(* IEC 61131-3 sources: SortJet_MasterSPS_Aufbau.fbsproj/09_Station/Stationen/_Basic/Aktionen, 11 files *)

(* ---- Basic_Shuttle_Aktion_FB_V01_00_00.fb.st ---- *)
(* METADATA
{
	"v3Meta": {
		"objectGuid": "f063b21c-ee9e-4ece-bc3c-2deffdcf07f3"
	}
}
*)
FUNCTION_BLOCK Basic_Shuttle_Aktion_FB_V01_00_00
VAR_IN_OUT

  // STRUKT
  BasisStationsParameter : StationBasisParameter_ST;

END_VAR
VAR_OUTPUT

  // BOOL
  bprtScheibe : BOOL;

END_VAR
VAR_INPUT

  // BOOL
  bpGeblaeseAktiv        : BOOL;
  bpAutomatikAktiv       : BOOL;
  bpVorAbAuftragAktiv    : BOOL;
  bpZielPositionErreicht : BOOL;

  // WORD
  wWand : WORD;

  // Bausteine
  Glastransport   : REFERENCE TO Shuttle_Glastransport_FB_V01_00_00;
  Kippen          : REFERENCE TO Shuttle_Kippen_V01_00_00;
  Wandverstellung : REFERENCE TO Dickenverstellung_FB_V01_00_00;
  Geblaese        : REFERENCE TO Geblaese_Schuetz_FB_V01_00_00;

END_VAR
VAR

  // Steps_TE
  steplAktion : STEPS_TE;

END_VAR
;
END_FUNCTION_BLOCK

(* ---- Basic_Station_Abnehmen_FB_V01_00_00.fb.st ---- *)
(* METADATA
{
	"v3Meta": {
		"objectGuid": "660d4460-1ddc-44b5-9e6a-0f9c596d74b5"
	}
}
*)
FUNCTION_BLOCK Basic_Station_Abnehmen_FB_V01_00_00 EXTENDS Basic_Station_Aktion_FB_V01_00_00
(* Hinweis:
   - Abnehmen: Station kippt, der Bediener nimmt die Scheiben ab und quittiert jede einzelne
   - Die Aktion schreibt nichts in den Glastransport
   - Kippen nur mit der Ausbaustufe bKippen
*)
VAR_INPUT

  // BOOLEAN
  bpFreigabeErhalten        : BOOL; // Station: Freigabe Si-Kreis (verzoegert) liegt an
  bpGlasAbgenommenQuittiert : BOOL; // Station: Bediener quittiert, dass die Scheibe abgenommen wurde (Taster oder Fusstaster gedrueckt)

  // Bausteine
  Kippen : REFERENCE TO Kippen_FB_V01_00_00;

END_VAR
VAR_OUTPUT

  // BOOLEAN
  bpAbnehmenLampe        : BOOL; // Ampel gruen
  bpSignalScheibeAbnehmen : BOOL; // Taster Scheibe abnehmen (blinkt)
  bpSignalGlasbruch      : BOOL;

END_VAR
VAR

  // INT
  ilScheibenZaehler : INT; // Anzahl der Scheiben, die noch abzunehmen sind

END_VAR
//-------------------------------------------------------------------------------------------------
// ABNEHMEN
//-------------------------------------------------------------------------------------------------
IF ( BasisStationsParameter.bAbnehmen
     AND bpAutomatikAktiv )
THEN
  (* Fehlerbehandlung:
     - Kippen
  *)
  IF ( Kippen.bpFehler ) THEN
    Kippen.bpPositionieren := FALSE;
    BasisStationsParameter.wFehlerNummer := Kippen.wpFehlerNr;
    steplAktion := STEP_900_E;
  END_IF

  CASE steplAktion OF
    // ABNEHMEN =====================
    STEP_0_E:
      (* Hinweis:
         - Freigabe durch Quittierten Si-Kreis da ?
      *)
      bpFehler := FALSE;
      bpSignalScheibeAbnehmen := FALSE;
      BasisStationsParameter.bAbnehmenAbgeschlossen := FALSE;

      IF ( bpFreigabeErhalten ) THEN
        ilScheibenZaehler := WORD_TO_INT( BasisStationsParameter.pAuftrag[cWAND_1].wAnzahlScheiben );
        steplAktion := STEP_10_E;
      END_IF

    // ABNEHMEN =====================
    STEP_10_E:
      (* Hinweis:
         - Pruefen ob das Geblase aktiv ist
           => Sicherung nicht ausgeloest
      *)
      IF ( bpGeblaeseFehler ) THEN
        bpDrosselklappeOeffnen := FALSE;
        BasisStationsParameter.wFehlerNummer := cMELDUNG_ANTRIEB_GEBLAESE;
        steplAktion := STEP_900_E;

      ELSE
        bpDrosselklappeOeffnen := TRUE;
        steplAktion := STEP_20_E;

      END_IF

    // ABNEHMEN =====================
    STEP_20_E:
      IF ( NOT Kippen.bpFehler ) THEN
        bpDrosselklappeOeffnen := TRUE;

        Kippen.epZielPosition := eKippen_Position_84Grad;
        Kippen.bpPositionieren := TRUE;

        steplAktion := STEP_30_E;
      ELSE
        Kippen.bpPositionieren := FALSE;
        BasisStationsParameter.wFehlerNummer := Kippen.wpFehlerNr;
        steplAktion := STEP_900_E;
      END_IF

    // ABNEHMEN =====================
    STEP_30_E:
      IF ( Kippen.bpDone OR NOT BasisStationsParameter.stMKs.stStationsAufbau.bKippen[cWAND_1] ) THEN
        bpDrosselklappeOeffnen := FALSE;
        Kippen.bpPositionieren := FALSE;

        bpAbnehmenLampe         := TRUE;
        bpSignalScheibeAbnehmen := TRUE;

        steplAktion := STEP_50_E;
      END_IF

    // ABNEHMEN =====================
    STEP_50_E:
      bpAbnehmenLampe         := gbFlashbit05sec;
      bpSignalScheibeAbnehmen := gbFlashbit05sec;

      (* Hinweis:
         - Erst die Lichtschranke unterbrechen und zur Station gehen
      *)
      IF ( bpFreigabeErhalten ) THEN
        steplAktion := STEP_60_E;
      END_IF

    // ABNEHMEN =====================
    STEP_60_E:
      bpAbnehmenLampe         := gbFlashbit05sec;
      bpSignalScheibeAbnehmen := gbFlashbit05sec;

      IF ( bpGlasAbgenommenQuittiert ) THEN
        ilScheibenZaehler := ( ilScheibenZaehler - 1 );

        IF ( ilScheibenZaehler > 0 ) THEN
          steplAktion := STEP_70_E;

        ELSE
          bpSignalGlasbruch       := FALSE;
          bpAbnehmenLampe         := FALSE;
          bpSignalScheibeAbnehmen := FALSE;

          steplAktion := STEP_1000_E;
        END_IF
      END_IF

    // ABNEHMEN =====================
    STEP_70_E:
      bpSignalGlasbruch := FALSE;

      IF ( NOT bpGlasAbgenommenQuittiert ) THEN
        steplAktion := STEP_60_E;
      END_IF

    // ABNEHMEN =====================
    STEP_900_E:
      bpFehler := TRUE;
      BasisStationsParameter.bFehler := TRUE;
      Kippen.bpPositionieren := FALSE;

    // ABNEHMEN =====================
    STEP_1000_E:
      BasisStationsParameter.bAbnehmenAbgeschlossen := TRUE;

  // ABNEHMEN =====================
  END_CASE
ELSE
  IF ( steplAktion > STEP_0_E ) THEN
    bpFehler                := FALSE;
    bpDrosselklappeOeffnen  := FALSE;
    bpSignalScheibeAbnehmen := FALSE;
    bpAbnehmenLampe         := FALSE;
    bpSignalGlasbruch       := FALSE;

    Kippen.bpPositionieren  := FALSE;

    BasisStationsParameter.bAbnehmenAbgeschlossen := FALSE;

    steplAktion := STEP_0_E;
  END_IF
END_IF
END_FUNCTION_BLOCK

(* ---- Basic_Station_Aktion_FB_V01_00_00.fb.st ---- *)
(* METADATA
{
	"v3Meta": {
		"objectGuid": "12c9ac0e-b17a-4793-9910-dd4830696017"
	}
}
*)
FUNCTION_BLOCK Basic_Station_Aktion_FB_V01_00_00
(* Hinweis:
   - Basis der wandweisen Aktionen einer Station (Ein-, Aus-, Durch-, Vortransport, Messkopplung)
   - Je Wand eine Instanz, die Station ruft sie in einer Schleife ueber die Waende auf
   - Die Komponenten (Kippen, Hub, Verstellungen ...) gibt es je Station nur einmal; die abgeleiteten
     Bausteine bekommen sie als Referenz
*)
VAR_IN_OUT

  // STRUKT
  BasisStationsParameter : StationBasisParameter_ST;

END_VAR
VAR_OUTPUT

  // BOOL
  bpFehler : BOOL; // Status: Schrittkette steht im Fehler
  bpDrosselklappeOeffnen : BOOL; // Anforderung an die Station: Drosselklappe oeffnen, solange der Transport laeuft (die Station entscheidet ueber den Ausgang)

END_VAR
VAR_INPUT

  // BOOL
  bpAutomatikAktiv       : BOOL;
  bpGeblaeseAktiv        : BOOL;
  bpGeblaeseFehler       : BOOL; // Station: Motorschutz des Geblaeses ausgeloest (Station ohne Geblaese-Baustein)
  bpZielPositionErreicht : BOOL;

  // WORD
  wWand : WORD;

  // Bausteine
  Glastransport : REFERENCE TO Basic_Glastransport_FB_V01_00_00;

END_VAR
VAR

  // Steps_TE
  steplAktion : STEPS_TE;

END_VAR
;
END_FUNCTION_BLOCK

(* ---- Basic_Station_Anlegen_FB_V01_00_00.fb.st ---- *)
(* METADATA
{
	"v3Meta": {
		"objectGuid": "7cf149bd-d1d2-4190-82d5-7daf21613ba4"
	}
}
*)
FUNCTION_BLOCK Basic_Station_Anlegen_FB_V01_00_00 EXTENDS Basic_Station_Aktion_FB_V01_00_00
(* Hinweis:
   - Anlegen von Hand: Die Hoehenkontrolle faehrt auf Position, ggf. Hubrahmen einfahren und Anschlaege ausfahren,
     dann wartet die Aktion auf die Quittierung des Bedieners (Taster / Fusstaster)
   - Die Aktion schreibt nichts in den Glastransport und liest nur die Sensoren
   - Ob angelegt oder eingetragen wird, entscheidet das MMI ueber die Transferstation des Auftrags
     (Transferstation 1 = eigene Station: Anlegen, Fremdanlage: Eintransport; Anlegetisch hinter einer Brechanlage)
   - Mit der VSG-Schnittstelle entscheidet die Station selbst: die Station (Eintransport Schneidlinie) uebernimmt ueber
     bpUebernahmeEintransport oder beendet das Anlegen ueber bpBetriebBeendet
   - Hubrahmen und Anschlag nur mit den Ausbaustufen bHubrahmen und bAnschlag, sonst muessen sie nicht uebergeben werden
*)
VAR_IN_OUT

  // BOOLEAN
  blAnlegenErzwingen : BOOL; // Anlegen wurde erzwungen, die Aktion nimmt die Anforderung entgegen

END_VAR
VAR_INPUT

  // BOOLEAN
  bpAnlegenQuittiert          : BOOL;        // Bediener hat angelegt (steigende Flanke Taster / Fusstaster)
  bpVoraussetzungErfuellt     : BOOL := TRUE; // Station: Voraussetzung zum Start (z.B. Kipparme frei)
  bpAnschlagAutomatischFahren : BOOL;        // Station: Anschlaege fahren automatisch aus
  bpNeustart                  : BOOL;        // Station: Anlegen von vorne beginnen (z.B. nach Umschalten der Anschlaege)
  bpUebernahmeEintransport    : BOOL;        // Station (VSG-Schnittstelle): Eintransport der Schneidlinie uebernimmt, das Anlegen gibt ab
  bpBetriebBeendet            : BOOL;        // Station (VSG-Schnittstelle): Automatikbetrieb der Schneidlinie beendet, Scheibe muss neu angelegt werden

  // Bausteine
  Messachse : REFERENCE TO Messachse_FB_V01_00_00;
  Anschlag  : REFERENCE TO ZylinderPneumatik_Anschlag_FB_V01_00_00;
  Hubrahmen : REFERENCE TO ZylinderPneumatik_Riemen_FB_V01_00_00;

END_VAR
VAR_OUTPUT

  // BOOLEAN
  bpAnlegenLampe          : BOOL; // Ampel gruen / Signal Scheibe aufgegeben (blinkt, bis angelegt ist)
  bpBedienerEingriff      : BOOL; // Aktion wartet auf den Bediener, Handfunktionen (Knebel, Hubrahmen) muessen im Automatikbetrieb greifen
  bpAnlegenInVorbereitung : BOOL; // Aktion fuehrt die Vorbereitung durch (vor dem Warten auf den Bediener)
  bpAnlegenAktiv          : BOOL; // Aktion ist gestartet und noch nicht abgeschlossen
  bpAnlegenFertig         : BOOL; // Aktion hat selbst abgeschlossen (epTypeHoehenmessung gueltig)
  bpGeblaeseAnforderung   : BOOL; // Geblaese soll laufen (Vorbereitung)
  bpGeblaeseStartenSensor : BOOL; // Der Einlaufsensor darf das Geblaese starten

  // TIME
  tpZeitBereitAnzulegen   : TIME; // Zeitpunkt, ab dem die Station bereit zum Anlegen ist (Statistik)

  // ENUM
  epTypeHoehenmessung     : ModusHoehenvermessung_EN;

END_VAR
VAR

  // BOOLEAN
  blAnschlagFehler       : BOOL;
  blAnschlagAusgefahren  : BOOL; // Anschlag ausgefahren oder nicht vorhanden
  blAnschlagFertig       : BOOL; // Anschlag fertig oder nicht vorhanden
  blHubrahmenFehler      : BOOL;
  blHubrahmenEingefahren : BOOL; // Hubrahmen eingefahren oder nicht vorhanden
  blSensorAnlegeseite    : BOOL; // Scheibe liegt an (Einlaufsensor belegt, Auslaufsensor frei)
  blSensorAuslaufBelegt  : BOOL;
  blModellscheibe        : BOOL;

END_VAR
//-------------------------------------------------------------------------------------------------
// ANLEGEN
//-------------------------------------------------------------------------------------------------
blAnschlagFehler       := FALSE;
blAnschlagAusgefahren  := TRUE;
blAnschlagFertig       := TRUE;
blHubrahmenFehler      := FALSE;
blHubrahmenEingefahren := TRUE;

IF ( BasisStationsParameter.stMKs.stStationsAufbau.bAnschlag ) THEN
  blAnschlagFehler      := Anschlag.bpFehler;
  blAnschlagAusgefahren := ( Anschlag.epStatusZylinder = eZylinderAusgefahren ) OR NOT bpAnschlagAutomatischFahren;
  blAnschlagFertig      := Anschlag.bpDone;
END_IF

IF ( BasisStationsParameter.stMKs.stStationsAufbau.bHubrahmen ) THEN
  blHubrahmenFehler      := Hubrahmen.bpFehler;
  blHubrahmenEingefahren := ( Hubrahmen.epStatusZylinder = eZylinderEingefahren );
END_IF

// Scheibe liegt an: Einlaufsensor belegt, auf der Gegenseite frei (mit Vorab-Sensor, wenn die Station damit misst)
IF ( BasisStationsParameter.stMKs.stStationsOptionen.stGlastransport.bScheibenmessungSensorVorabAuslauf ) THEN
  blSensorAuslaufBelegt := Glastransport.bpSensorAuslaufVorAb;
ELSE
  blSensorAuslaufBelegt := Glastransport.bpSensorAuslauf;
END_IF
blSensorAnlegeseite := Glastransport.bpSensorEinlauf AND NOT blSensorAuslaufBelegt;

blModellscheibe := ( BasisStationsParameter.wGlastyp[cWAND_1] = eScheibe_Modell );

IF( BasisStationsParameter.bAnlegen
    AND NOT BasisStationsParameter.bEintransport[cWAND_1]
    AND bpAutomatikAktiv )
THEN

  bpAnlegenAktiv := TRUE;

  // Ausnahmesituation
  IF ( BasisStationsParameter.stMKs.stStationsAufbau.bAnschlag ) THEN
    IF ( blAnschlagFehler ) THEN
      Anschlag.bpStartAusfahren := FALSE;
      Anschlag.bpStartEinfahren := FALSE;
      BasisStationsParameter.awFehlerInformationen[1] := cZYLINDER_ANSCHLAG;
      BasisStationsParameter.wFehlerNummer := Anschlag.wpFehlerNr;
      steplAktion := STEP_900_E;
    END_IF
  END_IF

  IF ( BasisStationsParameter.stMKs.stStationsAufbau.bHubrahmen ) THEN
    IF ( blHubrahmenFehler ) THEN
      Hubrahmen.bpStartAusfahren := FALSE;
      Hubrahmen.bpStartEinfahren := FALSE;
      BasisStationsParameter.awFehlerInformationen[1] := cZYLINDER_HUBRAHMEN;
      BasisStationsParameter.wFehlerNummer := Hubrahmen.wpFehlerNr;
      steplAktion := STEP_900_E;
    END_IF
  END_IF

  IF ( Messachse.bpFehler ) THEN
    Messachse.bpPositionierung := FALSE;
    BasisStationsParameter.wFehlerNummer := Messachse.wpFehlerNr;
    steplAktion := STEP_900_E;
  END_IF

  IF ( bpNeustart ) THEN
    steplAktion := STEP_0_E;
  END_IF

  CASE steplAktion OF
    // ANLEGEN ==================================
    STEP_0_E:
      (* Hinweis:
         - Variablen initalisieren
         - Starten des Anlegevorgangs
         - Voraussetzung der Station muss erfuellt sein, der Motorschutz des Geblaeses muss in Ordnung sein
      *)
      bpFehler                := FALSE;
      bpGeblaeseStartenSensor := FALSE;

      // Auftrag nach Status neu setzen. Bei Wiederholung (z.B. Messung fehlerhaft) will die Scheibe neu angelegt werden
      IF ( BasisStationsParameter.eStatusAuftrag = eAuftragWiederholen ) THEN
        BasisStationsParameter.eStatusAuftrag := eAuftragAktivWiederholen;
      ELSE
        BasisStationsParameter.eStatusAuftrag := eAuftragAktiv;
      END_IF

      IF ( bpGeblaeseFehler ) THEN
        BasisStationsParameter.wFehlerNummer := cMELDUNG_ANTRIEB_GEBLAESE;
        steplAktion := STEP_900_E;

      ELSIF ( bpVoraussetzungErfuellt ) THEN
        bpAnlegenLampe := FALSE;

        IF ( BasisStationsParameter.stMKs.stStationsAufbau.bAnschlag ) THEN
          Anschlag.bpStartEinfahren := FALSE;
          Anschlag.bpStartAusfahren := FALSE;
        END_IF

        IF ( bpUebernahmeEintransport ) THEN
          steplAktion := STEP_200_E;
        ELSE
          blAnlegenErzwingen := FALSE;
          steplAktion := STEP_10_E;
        END_IF

      END_IF

    // ANLEGEN ==============================
    STEP_10_E:
      (* Hinweis:
         - Hubrahmen einfahren sofern er es nicht ist
         - Anschlag Ausfahren sofern gefordert
         - Hoehenkontrolle auf Position fahren
      *)
      IF ( BasisStationsParameter.stMKs.stStationsAufbau.bHubrahmen ) THEN
        Hubrahmen.bpStartEinfahren := NOT blHubrahmenEingefahren;
      END_IF

      IF ( BasisStationsParameter.stMKs.stStationsAufbau.bAnschlag ) THEN
        Anschlag.bpStartAusfahren := bpAnschlagAutomatischFahren;
      END_IF

      IF ( BasisStationsParameter.stMKs.stStationsOptionen.stGlastransport.bScheibenVermessen ) THEN
        IF ( Messachse.Antrieb.rpMaxPosition < ( BasisStationsParameter.pAuftrag[cWAND_1].rAuftragsHoehe + Messachse.ppParameterBaustein.rKorrekturOffset ) ) THEN
          Messachse.rpZielPosition := Messachse.Antrieb.rpMaxPosition;
        ELSE
          Messachse.rpZielPosition := ( BasisStationsParameter.pAuftrag[cWAND_1].rAuftragsHoehe + Messachse.ppParameterBaustein.rKorrekturOffset );
        END_IF
      ELSE
        Messachse.rpZielPosition := BasisStationsParameter.stMKs.stGlasdaten[cWAND_1].rlMinGlasHoehe;
      END_IF
      Messachse.bpPositionierung := TRUE;

      steplAktion := STEP_20_E;

    // ANLEGEN ==============================
    STEP_20_E:
      (* Anmerkung:
         - Korrekte Stati der Zylinder und Achsen abfragen
         - Das Geblaese laeuft in der Vorbereitung
      *)
      bpGeblaeseAnforderung := TRUE;

      IF (     blHubrahmenEingefahren
           AND blAnschlagAusgefahren
           AND ( Messachse.bpDone OR NOT BasisStationsParameter.stMKs.stStationsOptionen.stGlastransport.bScheibenVermessen ) )
      THEN
        IF ( BasisStationsParameter.stMKs.stStationsAufbau.bHubrahmen ) THEN
          Hubrahmen.bpStartEinfahren := FALSE;
        END_IF

        IF ( BasisStationsParameter.stMKs.stStationsAufbau.bAnschlag ) THEN
          Anschlag.bpStartAusfahren := FALSE;
        END_IF

        Messachse.bpPositionierung := FALSE;
        bpGeblaeseAnforderung      := FALSE;

        // Anschlaege fahren nicht automatisch aus: erst auf den Taster warten, sonst direkt anlegen
        IF ( BasisStationsParameter.stMKs.stStationsAufbau.bAnschlag AND NOT bpAnschlagAutomatischFahren ) THEN
          steplAktion := STEP_30_E;
        ELSE
          tpZeitBereitAnzulegen  := TIME();
          bpDrosselklappeOeffnen := TRUE;
          steplAktion := STEP_100_E;
        END_IF

      END_IF

    // ANLEGEN ==============================
    STEP_30_E:
      (* Anmerkung:
         - Anschlaege fahren nicht automatisch aus, der Bediener faehrt sie mit dem Taster aus
         - Handfunktionen (Knebel, Hubrahmen) greifen im Automatikbetrieb
      *)
      bpAnlegenLampe := gbFlashbit05sec;

      // VSG-Schnittstelle: Automatikbetrieb beendet bzw. Eintransport wird uebernommen
      IF ( bpBetriebBeendet ) THEN
        BasisStationsParameter.eStatusAuftrag := eAuftragWiederholen;
        bpAnlegenLampe := FALSE;
        steplAktion := STEP_1000_E;
      END_IF

      IF ( bpUebernahmeEintransport ) THEN
        steplAktion := STEP_200_E;
      END_IF

      IF ( bpAnlegenQuittiert ) THEN
        Anschlag.bpStartAusfahren := TRUE;
        bpAnlegenLampe := FALSE;
        steplAktion := STEP_40_E;
      END_IF

      IF ( BasisStationsParameter.stMKs.stStationsAufbau.bHubrahmen ) THEN
        IF ( blHubrahmenFehler ) THEN
          Hubrahmen.bpStartEinfahren := FALSE;
          Hubrahmen.bpStartAusfahren := FALSE;

          BasisStationsParameter.awFehlerInformationen[1] := cZYLINDER_HUBRAHMEN;
          BasisStationsParameter.wFehlerNummer := Hubrahmen.wpFehlerNr;

          steplAktion := STEP_900_E;
        END_IF
      END_IF

    // ANLEGEN ==============================
    STEP_40_E:
      (* Anmerkung:
         - Anschlaege ausfahren
      *)
      IF ( blAnschlagFertig
           AND blAnschlagAusgefahren )
      THEN
        tpZeitBereitAnzulegen := TIME();

        Anschlag.bpStartAusfahren := FALSE;

        bpDrosselklappeOeffnen  := TRUE;
        bpAnlegenLampe          := TRUE;
        bpGeblaeseStartenSensor := TRUE;

        steplAktion := STEP_100_E;
      END_IF

    // ANLEGEN ==============================
    STEP_100_E:
      (* Anmerkung:
         - Warten bis der Bediener die Scheibe angelegt und quittiert hat
         - Geblaese starten wenn dieses nicht schon gestartet ist
           => Belegen des Einlaufsensors
         - Handfunktionen (Knebel, Hubrahmen) greifen im Automatikbetrieb
      *)
      IF ( blSensorAnlegeseite
           OR blModellscheibe )
      THEN
        bpAnlegenLampe := TRUE;
      ELSE
        bpAnlegenLampe := gbFlashbit05sec;
      END_IF

      bpGeblaeseStartenSensor := TRUE;

      // VSG-Schnittstelle: Automatikbetrieb beendet bzw. Eintransport wird uebernommen
      IF ( bpBetriebBeendet ) THEN
        BasisStationsParameter.eStatusAuftrag := eAuftragWiederholen;
        bpAnlegenLampe := FALSE;
        steplAktion := STEP_1000_E;
      END_IF

      IF ( bpUebernahmeEintransport ) THEN
        steplAktion := STEP_200_E;
      END_IF

      // Scheibe wurde angelegt
      IF ( bpAnlegenQuittiert
           AND ( blSensorAnlegeseite
                 OR blModellscheibe ) )
      THEN
        bpAnlegenLampe          := FALSE;
        bpGeblaeseStartenSensor := FALSE;

        BasisStationsParameter.dwWartezeit[cWAND_1] := TIME_TO_DWORD( TIME() - tpZeitBereitAnzulegen );

        bpDrosselklappeOeffnen := FALSE;

        BasisStationsParameter.eStatusAuftrag := eAuftragErfolgreich;

        // Wenn Modellscheibe -> Anschlaege einfahren
        IF ( blModellscheibe
             AND BasisStationsParameter.stMKs.stStationsAufbau.bAnschlag )
        THEN
          Anschlag.bpStartEinfahren := TRUE;
          Anschlag.bpStartAusfahren := FALSE;
          steplAktion := STEP_300_E;
        ELSE
          steplAktion := STEP_1000_E;
        END_IF

      END_IF

      (* Hinweis:
         - Der Auslauf- Sensor muss frei sein, um mit dem Einschleusen des Glases zu beginnen
      *)
      IF ( blSensorAuslaufBelegt
           AND bpAnlegenQuittiert
           AND NOT blModellscheibe )
      THEN
        wpgFehlerdaten[0] := BasisStationsParameter.stMKs.stStationsNummern.NummerExtern;
        SpsHinweis( eFehler_Station,
                    cMELDUNG_ANLEGEN_SENSOR_AUSLAUF_BELEGT,
                    BasisStationsParameter.stMKs.stStationsNummern.NummerIntern,
                    AutomatikkreisBestimmen( BasisStationsParameter.stMKs.stStationsNummern.NummerSPS ),
                    wpgFehlerdaten );
      END_IF

      (* Hinweis:
         - Der Einlaufsensor muss belegt sein
      *)
      IF ( NOT Glastransport.bpSensorEinlauf
           AND bpAnlegenQuittiert
           AND NOT blModellscheibe )
      THEN
        wpgFehlerdaten[0] := BasisStationsParameter.stMKs.stStationsNummern.NummerExtern;
        SpsHinweis( eFehler_Station,
                    cMELDUNG_ANLEGEN_SENSOR_EINLAUF_NICHT_BELEGT,
                    BasisStationsParameter.stMKs.stStationsNummern.NummerIntern,
                    AutomatikkreisBestimmen( BasisStationsParameter.stMKs.stStationsNummern.NummerSPS ),
                    wpgFehlerdaten );
      END_IF

      (* Fehlerbehandlung:
         - Hubpalette senkt / hebt nicht in der vorgeschriebenen Zeit bzw. Sensor schaltet nicht
      *)
      IF ( BasisStationsParameter.stMKs.stStationsAufbau.bHubrahmen ) THEN
        IF ( blHubrahmenFehler ) THEN
          Hubrahmen.bpStartEinfahren := FALSE;
          Hubrahmen.bpStartAusfahren := FALSE;

          BasisStationsParameter.awFehlerInformationen[1] := cZYLINDER_HUBRAHMEN;
          BasisStationsParameter.wFehlerNummer := Hubrahmen.wpFehlerNr;

          steplAktion := STEP_900_E;
        END_IF
      END_IF

    // ANLEGEN ==================================
    STEP_200_E:
      (* Anmerkung:
         - Die Station (Eintransport Schneidlinie) hat uebernommen: Glastransport, Hubrahmen, Anschlaege und
           Hoehenkontrolle gehoeren jetzt der Station, das Anlegen wartet bis der Auftrag beendet ist
      *)
      bpAnlegenLampe := FALSE;

    // ANLEGEN ==================================
    STEP_300_E:
      (* Anmerkung:
         - Anschlaege gesenkt
      *)
      IF ( blAnschlagFertig ) THEN
        Anschlag.bpStartEinfahren := FALSE;

        steplAktion := STEP_1000_E;
      END_IF

    // ANLEGEN ==================================
    STEP_900_E:
      BasisStationsParameter.eStatusAuftrag := eAuftragFehler;

      bpFehler := TRUE;
      BasisStationsParameter.bFehler := TRUE;

    // ANLEGEN ==================================
    STEP_1000_E:
      epTypeHoehenmessung := Modus_Positionieren_Auf_Oberkante_2_Sensoren;
      bpAnlegenFertig     := TRUE;

      BasisStationsParameter.bAnlegenAbgeschlossen := TRUE;

  // ANLEGEN ==================================
  END_CASE

  (* Hinweis:
     - Ausgaenge fuer die Station: Bediener-Eingriff (Handfunktionen im Automatikbetrieb) und Vorbereitung
  *)
  bpBedienerEingriff      := ( steplAktion = STEP_30_E ) OR ( steplAktion = STEP_100_E );
  bpAnlegenInVorbereitung := ( steplAktion <= STEP_20_E );
  bpAnlegenAktiv          := ( steplAktion <= STEP_100_E );

ELSE

  bpBedienerEingriff      := FALSE;
  bpAnlegenInVorbereitung := FALSE;
  bpAnlegenAktiv          := FALSE;

  IF( steplAktion > STEP_0_E ) THEN

    BasisStationsParameter.bAnlegenAbgeschlossen := FALSE;
    bpFehler                     := FALSE;
    bpAnlegenFertig              := FALSE;
    bpAnlegenLampe               := FALSE;
    bpGeblaeseAnforderung        := FALSE;
    bpGeblaeseStartenSensor      := FALSE;
    bpDrosselklappeOeffnen       := FALSE;
    Messachse.bpPositionierung   := FALSE;

    steplAktion := STEP_0_E;
  END_IF

END_IF
END_FUNCTION_BLOCK

(* ---- Basic_Station_Austransport_FB_V01_00_00.fb.st ---- *)
(* METADATA
{
	"v3Meta": {
		"objectGuid": "281ccc1c-3965-40cf-8682-0228b96383da"
	}
}
*)
FUNCTION_BLOCK Basic_Station_Austransport_FB_V01_00_00 EXTENDS Basic_Station_Aktion_FB_V01_00_00
VAR_INPUT

  // Bausteine
  Kippen          : REFERENCE TO Kippen_FB_V01_00_00;
  Hub             : REFERENCE TO Hub_FB_V01_00_00;
  Geblaese        : REFERENCE TO Geblaese_Schuetz_FB_V01_00_00;

  (* Hinweis:
     - Nur mit der Ausbaustufe bMessachse wird die Referenz benutzt,
       ohne diese Ausbaustufe muss die Station sie nicht uebergeben
  *)
  Messachse       : REFERENCE TO Messachse_FB_V01_00_00;

  (* Hinweis:
     - Nur mit der Ausbaustufe bDurchlaufSperreZumNachfolger wird die Referenz benutzt,
       ohne diese Ausbaustufe muss die Station sie nicht uebergeben
  *)
  Abschrankung      : REFERENCE TO ZylinderPneumatik_FB_V01_00_00;

END_VAR
VAR

  // BOOLEAN
  blQuelleWandLeer        : BOOL; // Auftrag: die Quellstation ist nach dem Austransport leer
  blVortransportGestartet : BOOL; // Vortransport vor dem Austransport (Option der Station) laeuft gemeinsam mit den Vorbewegungen
  blMessachseFertig       : BOOL; // Messachse auf Position oder nicht vorhanden
  blMitAbschrankung       : BOOL; // Austransport zum Nachfolger durch die bewegliche Abschrankung
  blAbschrankungFertig    : BOOL; // Abschrankung in der Endlage oder nicht beteiligt

END_VAR
//-------------------------------------------------------------------------------------------------
// AUSTRANSPORT
//-------------------------------------------------------------------------------------------------
blQuelleWandLeer := BasisStationsParameter.pAuftrag[wWand].stAuftragsInformationen.cBIT_SRCSTATION_EMPTY;
blMitAbschrankung := (     BasisStationsParameter.stMKs.stStationsAufbau.bDurchlaufSperreZumNachfolger
                       AND NOT BasisStationsParameter.bRueckwaertsTransportieren[wWand] );

IF ( BasisStationsParameter.bAustransport[wWand]
     AND bpAutomatikAktiv )
THEN

  // Ausnahmesituation
  IF ( Glastransport.bpFehler ) THEN
    Glastransport.bpAustransport             := FALSE;
    Glastransport.bpAustransportRueckwaertig := FALSE;
    Glastransport.bpVortransport             := FALSE;
    Glastransport.bpVortransportRueckwaertig := FALSE;
    Glastransport.bpReferenz                 := FALSE;
    bpDrosselklappeOeffnen                   := FALSE;
    BasisStationsParameter.wFehlerNummer := Glastransport.wpFehlerNr;
    steplAktion := STEP_900_E;
  END_IF

  IF ( Kippen.bpFehler ) THEN
    Kippen.bpPositionieren := FALSE;
    BasisStationsParameter.wFehlerNummer := Kippen.wpFehlerNr;
    steplAktion := STEP_900_E;
  END_IF

  IF ( Hub.bpFehler ) THEN
    Hub.bpStartHubAuf := FALSE;
    Hub.bpStartHubAb  := FALSE;
    BasisStationsParameter.wFehlerNummer := Hub.wpFehlerNr;
    steplAktion := STEP_900_E;
  END_IF

  IF ( bpGeblaeseFehler ) THEN
    BasisStationsParameter.wFehlerNummer := cMELDUNG_ANTRIEB_GEBLAESE;
    steplAktion := STEP_900_E;
  END_IF

  IF ( Geblaese.bpFehler )THEN
    BasisStationsParameter.wFehlerNummer := cMELDUNG_ANTRIEB_GEBLAESE;
    steplAktion := STEP_900_E;
  END_IF

  IF ( BasisStationsParameter.stMKs.stStationsAufbau.bMessachse ) THEN
    IF ( Messachse.bpFehler ) THEN
      Messachse.bpPositionierung := FALSE;
      BasisStationsParameter.wFehlerNummer := Messachse.wpFehlerNr;
      steplAktion := STEP_900_E;
    END_IF
  END_IF

  IF ( blMitAbschrankung ) THEN
    IF ( Abschrankung.bpFehler ) THEN
      Abschrankung.bpStartEinfahren := FALSE;
      Abschrankung.bpStartAusfahren := FALSE;
      BasisStationsParameter.awFehlerInformationen[1] := cZYLINDER_ABSCHRANKUNG;
      BasisStationsParameter.wFehlerNummer := Abschrankung.wpFehlerNr;
      steplAktion := STEP_900_E;
    END_IF
  END_IF

  CASE steplAktion OF
    // AUSTRANSPORT =====================
    STEP_0_E:
      (* Hinweis:
         - Geblaese aktiv und die Querfahrt hat die Zielposition erreicht (ohne Querfahrt immer erreicht)
      *)
      bpFehler := FALSE;
      blVortransportGestartet := FALSE;

      IF ( bpGeblaeseAktiv
           AND bpZielPositionErreicht )
      THEN
        Kippen.bpPositionieren := FALSE;
        bpDrosselklappeOeffnen := TRUE;

        steplAktion := STEP_10_E;
      END_IF

    // AUSTRANSPORT =====================
    STEP_10_E:
      (* Hinweis:
         - Ansteuerung Kippen
         - Hub auf die Sollposition des Auftrags fahren (nur Oben / Unten, sonst keine Bewegung)
         - Messachse auf die Auftragshoehe fahren (maximal bis zur Maximalposition)
         - Vortransport (Option der Station): Scheibe vor dem Austransport positionieren,
           laeuft gemeinsam mit den Bewegungen
      *)
      Kippen.epZielPosition  := BasisStationsParameter.pAuftrag[wWand].stAuftragsOptionen.eKippen_SollPosition;
      Kippen.bpPositionieren := TRUE;

      IF ( BasisStationsParameter.stMKs.stStationsAufbau.bHub ) THEN
        Hub.bpStartHubAuf := ( BasisStationsParameter.pAuftrag[wWand].stAuftragsOptionen.eHub = eHub_Oben );
        Hub.bpStartHubAb  := ( BasisStationsParameter.pAuftrag[wWand].stAuftragsOptionen.eHub = eHub_Unten );
      END_IF

      IF ( BasisStationsParameter.stMKs.stStationsAufbau.bMessachse ) THEN
        IF ( ( BasisStationsParameter.pAuftrag[wWand].rAuftragsHoehe + Messachse.ppParameterBaustein.rKorrekturOffset ) >= Messachse.Antrieb.rpMaxPosition ) THEN
          Messachse.rpZielPosition := Messachse.Antrieb.rpMaxPosition;
        ELSE
          Messachse.rpZielPosition := BasisStationsParameter.pAuftrag[wWand].rAuftragsHoehe + Messachse.ppParameterBaustein.rKorrekturOffset;
        END_IF
        Messachse.bpPositionierung := TRUE;
      END_IF

      blVortransportGestartet := BasisStationsParameter.stMKs.stStationsOptionen.stGlastransport.bVortransport;
      Glastransport.pAuftrag                   := BasisStationsParameter.pAuftrag[wWand];
      Glastransport.bpVortransport             := blVortransportGestartet AND NOT BasisStationsParameter.bRueckwaertsTransportieren[wWand];
      Glastransport.bpVortransportRueckwaertig := blVortransportGestartet AND     BasisStationsParameter.bRueckwaertsTransportieren[wWand];

      steplAktion := STEP_20_E;

    // AUSTRANSPORT =====================
    STEP_20_E:
      (* Hinweis:
         - Warten bis die Bewegungen und der Vortransport fertig sind
         - Der Vortransport wird abgebrochen, sobald der Empfaenger bereit zum Eintransport ist
      *)
      blMessachseFertig := TRUE;

      IF ( BasisStationsParameter.stMKs.stStationsAufbau.bMessachse ) THEN
        blMessachseFertig := Messachse.bpDone;
      END_IF

      (* Hinweis:
         - Bewegliche Abschrankung zum Nachfolger erst oeffnen (einfahren), wenn der Nachfolger bereit zum Eintransport ist
           (z.B. Drehstation steht in der Zielposition), vorher bleibt sie geschlossen
      *)
      blAbschrankungFertig := TRUE;

      IF ( blMitAbschrankung ) THEN
        // Erst auswerten, dann Kommando setzen: ein altes bpDone darf im Zyklus des Startens nicht als fertig zaehlen
        blAbschrankungFertig := ( Abschrankung.bpStartEinfahren AND Abschrankung.bpDone );

        IF ( BasisStationsParameter.InGlasTransportNachfolger[wWand].bBereitZumEintransport ) THEN
          Abschrankung.bpStartAusfahren := FALSE;
          Abschrankung.bpStartEinfahren := TRUE;
        END_IF
      END_IF

      Glastransport.bpAbbruchVortransport := blVortransportGestartet AND BasisStationsParameter.InGlasTransportNachfolger[wWand].bBereitZumEintransport;

      IF ( ( Kippen.bpDone OR NOT Kippen.bpPositionieren )
           AND blMessachseFertig
           AND blAbschrankungFertig
           AND ( Hub.bpDone OR NOT ( Hub.bpStartHubAuf OR Hub.bpStartHubAb ) OR NOT BasisStationsParameter.stMKs.stStationsAufbau.bHub )
           AND ( Glastransport.bpDone OR NOT blVortransportGestartet ) )
      THEN
        Kippen.bpPositionieren                   := FALSE;
        Hub.bpStartHubAuf                        := FALSE;
        Hub.bpStartHubAb                         := FALSE;
        Glastransport.bpAbbruchVortransport      := FALSE;
        Glastransport.bpVortransport             := FALSE;
        Glastransport.bpVortransportRueckwaertig := FALSE;
        blVortransportGestartet                  := FALSE;

        IF ( BasisStationsParameter.stMKs.stStationsAufbau.bMessachse ) THEN
          Messachse.bpPositionierung := FALSE;
        END_IF

        steplAktion := STEP_100_E;
      END_IF

    // AUSTRANSPORT =====================
    STEP_100_E:
      (* Hinweis:
         - Austransport starten
      *)
      Glastransport.pAuftrag := BasisStationsParameter.pAuftrag[wWand];
      Glastransport.bpAustransport             := BasisStationsParameter.bAustransport[wWand] AND NOT BasisStationsParameter.bRueckwaertsTransportieren[wWand];
      Glastransport.bpAustransportRueckwaertig := BasisStationsParameter.bAustransport[wWand] AND     BasisStationsParameter.bRueckwaertsTransportieren[wWand];

      steplAktion := STEP_110_E;

    // AUSTRANSPORT =====================
    STEP_110_E:
      (* Hinweis:
         - Bei letzter Scheibe und Station leer -> Kippen
      *)
      IF ( Glastransport.bpFreigabeFremdprozess
           AND BasisStationsParameter.pAuftrag[wWand].bLetzteScheibe
           AND blQuelleWandLeer )
      THEN
        Kippen.epZielPosition := BasisStationsParameter.pAuftrag[wWand].stAuftragsOptionen.eKippen_SollPosition_NachAustransport;
        Kippen.bpPositionieren := TRUE;

        IF ( BasisStationsParameter.stMKs.stStationsAufbau.bHub ) THEN
          Hub.bpStartHubAuf := ( BasisStationsParameter.pAuftrag[wWand].stAuftragsOptionen.eHub_NachAustransport = eHub_Oben );
          Hub.bpStartHubAb  := ( BasisStationsParameter.pAuftrag[wWand].stAuftragsOptionen.eHub_NachAustransport = eHub_Unten );
        END_IF
      END_IF

      (* Hinweis:
         - Austransport abgeschlossen
      *)
      IF ( Glastransport.bpDone ) THEN
        Glastransport.bpAustransport             := FALSE;
        Glastransport.bpAustransportRueckwaertig := FALSE;
        bpDrosselklappeOeffnen                   := FALSE;

        (* Hinweis:
           - Bewegliche Abschrankung zum Nachfolger schliessen (ausfahren)
        *)
        IF ( blMitAbschrankung ) THEN
          Abschrankung.bpStartEinfahren := FALSE;
          Abschrankung.bpStartAusfahren := TRUE;
        END_IF

        steplAktion := STEP_200_E;

      END_IF

    // AUSTRANSPORT =====================
    STEP_200_E:
      (* Hinweis:
         - Austransport ist vorbei: die Achsen des Glastransports abnullen (Zaehlerueberlauf des Gebers),
           ein Slave-Antrieb des eigenen Glastransports wird dabei vom Master abgekoppelt
         - Nur nach dem Austransport, nie im Eintransport
         - Bei letzter Scheibe und Station leer -> Kippen, gemeinsam mit dem Abnullen
      *)
      Glastransport.bpReferenz := TRUE;

      IF BasisStationsParameter.pAuftrag[wWand].bLetzteScheibe
         AND blQuelleWandLeer
      THEN
        Kippen.epZielPosition := BasisStationsParameter.pAuftrag[wWand].stAuftragsOptionen.eKippen_SollPosition_NachAustransport;
        Kippen.bpPositionieren := TRUE;

        (* Hinweis:
           - Hub auf die Sollposition nach dem Austransport fahren (nur Oben / Unten, sonst keine Bewegung)
        *)
        IF ( BasisStationsParameter.stMKs.stStationsAufbau.bHub ) THEN
          Hub.bpStartHubAuf := ( BasisStationsParameter.pAuftrag[wWand].stAuftragsOptionen.eHub_NachAustransport = eHub_Oben );
          Hub.bpStartHubAb  := ( BasisStationsParameter.pAuftrag[wWand].stAuftragsOptionen.eHub_NachAustransport = eHub_Unten );
        END_IF
      END_IF

      steplAktion := STEP_210_E;

    // AUSTRANSPORT =====================
    STEP_210_E:
      blAbschrankungFertig := TRUE;

      IF ( blMitAbschrankung ) THEN
        blAbschrankungFertig := Abschrankung.bpDone;
      END_IF

      IF ( ( Kippen.bpDone OR NOT Kippen.bpPositionieren )
           AND ( Hub.bpDone OR NOT ( Hub.bpStartHubAuf OR Hub.bpStartHubAb ) OR NOT BasisStationsParameter.stMKs.stStationsAufbau.bHub )
           AND Glastransport.bpDone
           AND blAbschrankungFertig )
      THEN
        Kippen.bpPositionieren   := FALSE;
        Hub.bpStartHubAuf        := FALSE;
        Hub.bpStartHubAb         := FALSE;
        Glastransport.bpReferenz := FALSE;

        IF ( blMitAbschrankung ) THEN
          Abschrankung.bpStartAusfahren := FALSE;
        END_IF

        steplAktion := STEP_1000_E;
      END_IF

    // AUSTRANSPORT =====================
    STEP_900_E:
      bpFehler := TRUE;
      BasisStationsParameter.bFehler := TRUE;

    // AUSTRANSPORT =====================
    STEP_1000_E:
      BasisStationsParameter.bAustransportAbgeschlossen[wWand] := TRUE;

  // AUSTRANSPORT =====================
  END_CASE
ELSE

  IF (steplAktion > STEP_0_E) THEN
    bpFehler := FALSE;
    bpDrosselklappeOeffnen := FALSE;
    BasisStationsParameter.bAustransportAbgeschlossen[wWand] := FALSE;

    Kippen.bpPositionieren                   := FALSE;
    Hub.bpStartHubAuf                        := FALSE;
    Hub.bpStartHubAb                         := FALSE;
    Glastransport.bpAustransport             := FALSE;
    Glastransport.bpAustransportRueckwaertig := FALSE;
    Glastransport.bpVortransport             := FALSE;
    Glastransport.bpVortransportRueckwaertig := FALSE;
    Glastransport.bpAbbruchVortransport      := FALSE;
    Glastransport.bpReferenz                 := FALSE;
    blVortransportGestartet                  := FALSE;

    IF ( BasisStationsParameter.stMKs.stStationsAufbau.bMessachse ) THEN
      Messachse.bpPositionierung := FALSE;
    END_IF

    IF ( BasisStationsParameter.stMKs.stStationsAufbau.bDurchlaufSperreZumNachfolger ) THEN
      Abschrankung.bpStartEinfahren := FALSE;
      Abschrankung.bpStartAusfahren := FALSE;
    END_IF

    steplAktion := STEP_0_E;
  END_IF

END_IF
END_FUNCTION_BLOCK

(* ---- Basic_Station_Durchtransport_FB_V01_00_00.fb.st ---- *)
(* METADATA
{
	"v3Meta": {
		"objectGuid": "ca80c58d-93c1-43cb-beb6-89c88c6be1a7"
	}
}
*)
FUNCTION_BLOCK Basic_Station_Durchtransport_FB_V01_00_00 EXTENDS Basic_Station_Aktion_FB_V01_00_00
VAR_INPUT

  // Bausteine
  Hub : REFERENCE TO Hub_FB_V01_00_00;

END_VAR
//-------------------------------------------------------------------------------------------------
// DURCHTRANSPORT
//-------------------------------------------------------------------------------------------------
IF ( BasisStationsParameter.bDurchtransport[wWand]
     AND bpAutomatikAktiv )
THEN

  // Ausnahmesituation
  IF ( Glastransport.bpFehler ) THEN
    Glastransport.bpDurchtransport := FALSE;
    BasisStationsParameter.wFehlerNummer := Glastransport.wpFehlerNr;
    steplAktion := STEP_900_E;
  END_IF

  IF ( Hub.bpFehler ) THEN
    Hub.bpStartHubAuf := FALSE;
    Hub.bpStartHubAb  := FALSE;
    BasisStationsParameter.wFehlerNummer := Hub.wpFehlerNr;
    steplAktion := STEP_900_E;
  END_IF

  CASE steplAktion OF
    // DURCHTRANSPORT =============================
    STEP_0_E:
      bpFehler := FALSE;
      BasisStationsParameter.bDurchtransportAbgeschlossen[wWand] := FALSE;

      steplAktion := STEP_5_E;

    // DURCHTRANSPORT =============================
    STEP_5_E:
      (* Hinweis:
         - Hub auf die Sollposition des Auftrags fahren (nur Oben / Unten, sonst keine Bewegung)
      *)
      IF ( BasisStationsParameter.stMKs.stStationsAufbau.bHub ) THEN
        Hub.bpStartHubAuf := ( BasisStationsParameter.pAuftrag[wWand].stAuftragsOptionen.eHub = eHub_Oben );
        Hub.bpStartHubAb  := ( BasisStationsParameter.pAuftrag[wWand].stAuftragsOptionen.eHub = eHub_Unten );
      END_IF

      steplAktion := STEP_6_E;

    // DURCHTRANSPORT =============================
    STEP_6_E:
      IF ( Hub.bpDone OR NOT ( Hub.bpStartHubAuf OR Hub.bpStartHubAb ) OR NOT BasisStationsParameter.stMKs.stStationsAufbau.bHub ) THEN
        Hub.bpStartHubAuf := FALSE;
        Hub.bpStartHubAb  := FALSE;
        steplAktion := STEP_10_E;
      END_IF

    // DURCHTRANSPORT =============================
    STEP_10_E:
      Glastransport.pAuftrag := BasisStationsParameter.pAuftrag[wWand];
      Glastransport.bpDurchtransport := TRUE;

      steplAktion := STEP_20_E;

    // DURCHTRANSPORT =============================
    STEP_20_E:
      IF ( Glastransport.bpDone )  THEN
        Glastransport.bpDurchtransport := FALSE;
        steplAktion := STEP_1000_E;
      END_IF

    // DURCHTRANSPORT =============================
    STEP_900_E:
      bpFehler := TRUE;
      BasisStationsParameter.bFehler := TRUE;

    // DURCHTRANSPORT =============================
    STEP_1000_E:
      BasisStationsParameter.bDurchtransportAbgeschlossen[wWand] := TRUE;

  // DURCHTRANSPORT =============================
  END_CASE
ELSE

  IF (steplAktion > STEP_0_E) THEN
    bpFehler := FALSE;
    BasisStationsParameter.bDurchtransportAbgeschlossen[wWand] := FALSE;
    Glastransport.bpDurchtransport := FALSE;
    Hub.bpStartHubAuf := FALSE;
    Hub.bpStartHubAb  := FALSE;

    steplAktion := STEP_0_E;
  END_IF

END_IF
END_FUNCTION_BLOCK

(* ---- Basic_Station_Eintransport_FB_V01_00_00.fb.st ---- *)
(* METADATA
{
	"v3Meta": {
		"objectGuid": "0e6ffebb-2f8e-4d3e-883f-b07758de8e3e"
	}
}
*)
FUNCTION_BLOCK Basic_Station_Eintransport_FB_V01_00_00 EXTENDS Basic_Station_Aktion_FB_V01_00_00
VAR_INPUT

  // Bausteine
  Kippen          : REFERENCE TO Kippen_FB_V01_00_00;
  Hub             : REFERENCE TO Hub_FB_V01_00_00;
  Roellchenleiste : REFERENCE TO ZylinderPneumatik_3Wege_FB_V01_00_00;
  Wandverstellung : REFERENCE TO ZylinderPneumatik_3Wege_FB_V01_00_00;
  Geblaese        : REFERENCE TO Geblaese_Schuetz_FB_V01_00_00;

  (* Hinweis:
     - Nur mit den Ausbaustufen bMessachse und bTransportVerstellung wird die Referenz benutzt,
       ohne diese Ausbaustufe muss die Station sie nicht uebergeben
  *)
  Messachse         : REFERENCE TO Messachse_FB_V01_00_00;
  Dickenverstellung : REFERENCE TO ZylinderPneumatik_3Wege_FB_V01_00_00;

  (* Hinweis:
     - Nur mit der Ausbaustufe bDurchlaufSperreZumNachfolger wird die Referenz benutzt,
       ohne diese Ausbaustufe muss die Station sie nicht uebergeben
  *)
  Abschrankung      : REFERENCE TO ZylinderPneumatik_FB_V01_00_00;

END_VAR
VAR

  // BOOLEAN
  blVortransportGestartet : BOOL; // Vortransport zum Vorab-Sensor laeuft gemeinsam mit den Nachbewegungen
  blMessachseFertig       : BOOL; // Messachse auf Position oder nicht vorhanden
  blDickenverstellungFertig : BOOL; // Dickenverstellung auf Position oder nicht vorhanden
  blMitAbschrankung         : BOOL; // Rueckwaertiger Eintransport vom Nachfolger durch die bewegliche Abschrankung
  blAbschrankungFertig      : BOOL; // Abschrankung in der Endlage oder nicht beteiligt

END_VAR
//-------------------------------------------------------------------------------------------------
// EINTRANSPORT
//-------------------------------------------------------------------------------------------------
blMitAbschrankung := (     BasisStationsParameter.stMKs.stStationsAufbau.bDurchlaufSperreZumNachfolger
                       AND BasisStationsParameter.bRueckwaertsTransportieren[wWand] );

IF ( BasisStationsParameter.bEintransport[wWand]
     AND bpAutomatikAktiv )
THEN

  // Ausnahmesituation
  IF ( Glastransport.bpFehler ) THEN
    Glastransport.bpEintransport             := FALSE;
    Glastransport.bpEintransportRueckwaertig := FALSE;
    Glastransport.bpVortransport             := FALSE;
    Glastransport.bpVortransportRueckwaertig := FALSE;
    bpDrosselklappeOeffnen                   := FALSE;
    BasisStationsParameter.wFehlerNummer := Glastransport.wpFehlerNr;
    steplAktion := STEP_900_E;
  END_IF

  IF ( Kippen.bpFehler ) THEN
    Kippen.bpPositionieren := FALSE;
    BasisStationsParameter.wFehlerNummer := Kippen.wpFehlerNr;
    steplAktion := STEP_900_E;
  END_IF

  IF ( Hub.bpFehler ) THEN
    Hub.bpStartHubAb  := FALSE;
    Hub.bpStartHubAuf := FALSE;
    BasisStationsParameter.wFehlerNummer := Hub.wpFehlerNr;
    steplAktion := STEP_900_E;
  END_IF

  IF ( Roellchenleiste.bpFehler ) THEN
    Roellchenleiste.bpStartPneumatik := FALSE;
    BasisStationsParameter.awFehlerInformationen[1] := cZYLINDER_ROELLCHENLEISTE;
    BasisStationsParameter.wFehlerNummer := Roellchenleiste.wpFehlerNr;
    steplAktion := STEP_900_E;
  END_IF

  IF ( Wandverstellung.bpFehler ) THEN
    Wandverstellung.bpStartPneumatik := FALSE;
    BasisStationsParameter.awFehlerInformationen[1] := cZYLINDER_WANDVERSTELLUNG;
    BasisStationsParameter.wFehlerNummer := Wandverstellung.wpFehlerNr;
    steplAktion := STEP_900_E;
  END_IF

  IF ( bpGeblaeseFehler ) THEN
    BasisStationsParameter.wFehlerNummer := cMELDUNG_ANTRIEB_GEBLAESE;
    steplAktion := STEP_900_E;
  END_IF

  IF ( Geblaese.bpFehler ) THEN
    BasisStationsParameter.wFehlerNummer := cMELDUNG_ANTRIEB_GEBLAESE;
    steplAktion := STEP_900_E;
  END_IF

  IF ( BasisStationsParameter.stMKs.stStationsAufbau.bMessachse ) THEN
    IF ( Messachse.bpFehler ) THEN
      Messachse.bpPositionierung := FALSE;
      BasisStationsParameter.wFehlerNummer := Messachse.wpFehlerNr;
      steplAktion := STEP_900_E;
    END_IF
  END_IF

  IF ( BasisStationsParameter.stMKs.stStationsAufbau.bTransportVerstellung[wWand] ) THEN
    IF ( Dickenverstellung.bpFehler ) THEN
      Dickenverstellung.bpStartPneumatik := FALSE;
      BasisStationsParameter.awFehlerInformationen[1] := cZYLINDER_DICKENVERSTELLUNG;
      BasisStationsParameter.wFehlerNummer := Dickenverstellung.wpFehlerNr;
      steplAktion := STEP_900_E;
    END_IF
  END_IF

  IF ( blMitAbschrankung ) THEN
    IF ( Abschrankung.bpFehler ) THEN
      Abschrankung.bpStartEinfahren := FALSE;
      Abschrankung.bpStartAusfahren := FALSE;
      BasisStationsParameter.awFehlerInformationen[1] := cZYLINDER_ABSCHRANKUNG;
      BasisStationsParameter.wFehlerNummer := Abschrankung.wpFehlerNr;
      steplAktion := STEP_900_E;
    END_IF
  END_IF

  CASE steplAktion OF
    // EINTRANSPORT ===============================
    STEP_0_E:
      (* Hinweis:
         - Variablen zuruecksetzen
      *)
      bpFehler := FALSE;
      blVortransportGestartet := FALSE;

      (* Hinweis:
         - Pruefen ob die Querfahrt die Zielposition erreicht hat (ohne Querfahrt immer erreicht)
      *)
      IF ( bpZielPositionErreicht ) THEN
        steplAktion := STEP_10_E;
      END_IF

    // EINTRANSPORT ===============================
    STEP_10_E:
      (* Hinweis:
         - Pruefen ob die Geblase aktiv sind
      *)
      IF ( bpGeblaeseAktiv ) THEN
        bpDrosselklappeOeffnen := TRUE;

        Roellchenleiste.epOeffnungsStellung := BasisStationsParameter.pAuftrag[wWand].stAuftragsOptionen.eDickenverstellung;
        Roellchenleiste.bpStartPneumatik := TRUE;

        Wandverstellung.epOeffnungsStellung := BasisStationsParameter.pAuftrag[wWand].stAuftragsOptionen.eDickenverstellung;
        Wandverstellung.bpStartPneumatik := TRUE;

        (* Hinweis:
           - Dickenverstellung nach der Glasdicke aus dem Auftrag (entschieden in der Basis-Schrittkette)
           - Messachse auf die Auftragshoehe fahren
        *)
        IF ( BasisStationsParameter.stMKs.stStationsAufbau.bTransportVerstellung[wWand] ) THEN
          Dickenverstellung.epOeffnungsStellung := BasisStationsParameter.pAuftrag[wWand].stAuftragsOptionen.eDickenverstellung;
          Dickenverstellung.bpStartPneumatik := TRUE;
        END_IF

        IF ( BasisStationsParameter.stMKs.stStationsAufbau.bMessachse ) THEN
          Messachse.rpZielPosition := BasisStationsParameter.pAuftrag[wWand].rAuftragsHoehe + Messachse.ppParameterBaustein.rKorrekturOffset;
          Messachse.bpPositionierung := TRUE;
        END_IF

        Kippen.epZielPosition := BasisStationsParameter.pAuftrag[wWand].stAuftragsOptionen.eKippen_SollPosition;
        Kippen.bpPositionieren := TRUE;

        (* Hinweis:
           - Hub auf die Sollposition des Auftrags fahren (nur Oben / Unten, sonst keine Bewegung)
        *)
        IF ( BasisStationsParameter.stMKs.stStationsAufbau.bHub ) THEN
          Hub.bpStartHubAuf := ( BasisStationsParameter.pAuftrag[wWand].stAuftragsOptionen.eHub = eHub_Oben );
          Hub.bpStartHubAb  := ( BasisStationsParameter.pAuftrag[wWand].stAuftragsOptionen.eHub = eHub_Unten );
        END_IF

        (* Hinweis:
           - Bewegliche Abschrankung zum Nachfolger oeffnen (einfahren)
        *)
        IF ( blMitAbschrankung ) THEN
          Abschrankung.bpStartAusfahren := FALSE;
          Abschrankung.bpStartEinfahren := TRUE;
        END_IF

        steplAktion := STEP_20_E;
      END_IF

    // EINTRANSPORT ===============================
    STEP_20_E:
      blMessachseFertig         := TRUE;
      blDickenverstellungFertig := TRUE;

      IF ( BasisStationsParameter.stMKs.stStationsAufbau.bMessachse ) THEN
        blMessachseFertig := Messachse.bpDone;
      END_IF

      IF ( BasisStationsParameter.stMKs.stStationsAufbau.bTransportVerstellung[wWand] ) THEN
        blDickenverstellungFertig := Dickenverstellung.bpDone;
      END_IF

      blAbschrankungFertig := TRUE;

      IF ( blMitAbschrankung ) THEN
        blAbschrankungFertig := Abschrankung.bpDone;
      END_IF

      IF ( ( Kippen.bpDone )
           AND blMessachseFertig
           AND blDickenverstellungFertig
           AND blAbschrankungFertig
           AND ( Roellchenleiste.bpDone OR NOT BasisStationsParameter.stMKs.stStationsAufbau.bRoellchenleiste[wWand] )
           AND ( Wandverstellung.bpDone OR NOT BasisStationsParameter.stMKs.stStationsAufbau.bWandverstellung[wWand] )
           AND ( Hub.bpDone OR NOT ( Hub.bpStartHubAuf OR Hub.bpStartHubAb ) OR NOT BasisStationsParameter.stMKs.stStationsAufbau.bHub ) )
      THEN
        Roellchenleiste.bpStartPneumatik := FALSE;
        Wandverstellung.bpStartPneumatik := FALSE;
        Kippen.bpPositionieren           := FALSE;
        Hub.bpStartHubAuf                := FALSE;
        Hub.bpStartHubAb                 := FALSE;

        IF ( BasisStationsParameter.stMKs.stStationsAufbau.bTransportVerstellung[wWand] ) THEN
          Dickenverstellung.bpStartPneumatik := FALSE;
        END_IF

        IF ( BasisStationsParameter.stMKs.stStationsAufbau.bMessachse ) THEN
          Messachse.bpPositionierung := FALSE;
        END_IF

        steplAktion := STEP_100_E;
      END_IF

    // EINTRANSPORT =====================
    STEP_100_E:
      // ---------------------------------------------------------------------------------------
      //  STARTEN DES EINTRANSPORTS
      //
      //  Hinweis:
      //  - n/c
      // ---------------------------------------------------------------------------------------
      Glastransport.eGlastyp                   := BasisStationsParameter.wGlasTyp[wWand];
      Glastransport.bpScheibentrennen          := BasisStationsParameter.bScheibentrennen[wWand];
      Glastransport.pAuftrag                   := BasisStationsParameter.pAuftrag[wWand];
      Glastransport.bpEintransport             := BasisStationsParameter.bEintransport[wWand] AND NOT BasisStationsParameter.bRueckwaertsTransportieren[wWand];
      Glastransport.bpEintransportRueckwaertig := BasisStationsParameter.bEintransport[wWand] AND     BasisStationsParameter.bRueckwaertsTransportieren[wWand];

      steplAktion := STEP_110_E;

    // EINTRANSPORT =====================
    STEP_110_E:
      IF  ( Glastransport.bpFreigabeFremdprozess
            AND BasisStationsParameter.pAuftrag[wWand].bLetzteScheibe )
      THEN
        (* Hinweis:
           - Richtung ist Invertiert zur Eintransport- Position
        *)
        Kippen.epZielPosition := BasisStationsParameter.pAuftrag[wWand].stAuftragsOptionen.eKippen_SollPosition_NachEintransport;
        Kippen.bpLangsamKippen := (     (    ( Kippen.epZielPosition = eKippen_Position_90Grad )
                                          OR ( Kippen.epZielPosition = eKippen_Position_84Grad ) )
                                    AND (    ( BasisStationsParameter.pAuftrag[wWand].rAuftragsDicke < 3 )
                                          OR ( BasisStationsParameter.pAuftrag[wWand].rAuftragsHoehe > 1200 ) ) );
        Kippen.bpPositionieren := TRUE;

        IF ( BasisStationsParameter.stMKs.stStationsAufbau.bHub ) THEN
          Hub.bpStartHubAuf := ( BasisStationsParameter.pAuftrag[wWand].stAuftragsOptionen.eHub_NachEintransport = eHub_Oben );
          Hub.bpStartHubAb  := ( BasisStationsParameter.pAuftrag[wWand].stAuftragsOptionen.eHub_NachEintransport = eHub_Unten );
        END_IF
      END_IF

      IF ( Glastransport.bpDone ) THEN
        Glastransport.bpEintransport             := FALSE;
        Glastransport.bpEintransportRueckwaertig := FALSE;
        bpDrosselklappeOeffnen                   := FALSE;

        (* Hinweis:
           - Bewegliche Abschrankung zum Nachfolger schliessen (ausfahren)
        *)
        IF ( blMitAbschrankung ) THEN
          Abschrankung.bpStartEinfahren := FALSE;
          Abschrankung.bpStartAusfahren := TRUE;
        END_IF

        steplAktion := STEP_150_E;
      END_IF

    // EINTRANSPORT =====================
    STEP_150_E:
      (* Hinweis:
         - Warten bis die bewegliche Abschrankung geschlossen ist (ohne Abschrankung sofort weiter)
      *)
      blAbschrankungFertig := TRUE;

      IF ( blMitAbschrankung ) THEN
        blAbschrankungFertig := Abschrankung.bpDone;
      END_IF

      IF ( blAbschrankungFertig ) THEN
        IF ( blMitAbschrankung ) THEN
          Abschrankung.bpStartAusfahren := FALSE;
        END_IF

        IF ( BasisStationsParameter.pAuftrag[wWand].bLetzteScheibe) THEN
          steplAktion := STEP_200_E;
        ELSE
          steplAktion := STEP_1000_E;
        END_IF
      END_IF

    // EINTRANSPORT =====================
    STEP_200_E:
      // ---------------------------------------------------------------------------------------
      //  OPTIONAL - KOMPONENTEN STEUERUNG
      //
      //  Hinweis:
      //  - Ausrichtung der Station fuer den Austransport
      //  - Der Vortransport zum Vorab-Sensor laeuft gleichzeitig mit den Nachbewegungen
      // ---------------------------------------------------------------------------------------

      (* Hinweis:
         - Richtung ist Invertiert zur Eintransport- Position
      *)
      Kippen.epZielPosition := BasisStationsParameter.pAuftrag[wWand].stAuftragsOptionen.eKippen_SollPosition_NachEintransport;
      Kippen.bpLangsamKippen := (     (    ( Kippen.epZielPosition = eKippen_Position_90Grad )
                                            OR ( Kippen.epZielPosition = eKippen_Position_84Grad ) )
                                  AND (    ( BasisStationsParameter.pAuftrag[wWand].rAuftragsDicke < 3 )
                                       OR ( BasisStationsParameter.pAuftrag[wWand].rAuftragsHoehe > 1200 ) ) );
      Kippen.bpPositionieren := TRUE;

      (* Hinweis:
         - Hub auf die Sollposition nach dem Eintransport fahren (nur Oben / Unten, sonst keine Bewegung)
      *)
      IF ( BasisStationsParameter.stMKs.stStationsAufbau.bHub ) THEN
        Hub.bpStartHubAuf := ( BasisStationsParameter.pAuftrag[wWand].stAuftragsOptionen.eHub_NachEintransport = eHub_Oben );
        Hub.bpStartHubAb  := ( BasisStationsParameter.pAuftrag[wWand].stAuftragsOptionen.eHub_NachEintransport = eHub_Unten );
      END_IF

      (* Hinweis:
         - Auslauf-Vorab (rueckwaerts Einlauf-Vorab): nach dem Sammeln positioniert der Vortransport die Scheibe auf den Vorab-Sensor
      *)
      blVortransportGestartet := (     (     NOT BasisStationsParameter.bRueckwaertsTransportieren[wWand]
                                         AND ( BasisStationsParameter.pAuftrag[wWand].stAuftragsOptionen.eGlastransport = eGlastransport_AufAuslaufVorab ) )
                                   OR  (     BasisStationsParameter.bRueckwaertsTransportieren[wWand]
                                         AND ( BasisStationsParameter.pAuftrag[wWand].stAuftragsOptionen.eGlastransport = eGlastransport_AufEinlaufVorab ) ) );
      Glastransport.bpVortransport             := blVortransportGestartet AND NOT BasisStationsParameter.bRueckwaertsTransportieren[wWand];
      Glastransport.bpVortransportRueckwaertig := blVortransportGestartet AND     BasisStationsParameter.bRueckwaertsTransportieren[wWand];

      steplAktion := STEP_210_E;

    // EINTRANSPORT =====================
    STEP_210_E:
      (* Hinweis:
         - Warten bis die Nachbewegungen und der Vortransport fertig sind
      *)
      IF ( ( Kippen.bpDone OR NOT Kippen.bpPositionieren )
           AND ( Hub.bpDone OR NOT ( Hub.bpStartHubAuf OR Hub.bpStartHubAb ) OR NOT BasisStationsParameter.stMKs.stStationsAufbau.bHub )
           AND ( Glastransport.bpDone OR NOT blVortransportGestartet ) )
      THEN
        Kippen.bpPositionieren                   := FALSE;
        Kippen.bpLangsamKippen                   := FALSE;
        Hub.bpStartHubAuf                        := FALSE;
        Hub.bpStartHubAb                         := FALSE;
        Glastransport.bpVortransport             := FALSE;
        Glastransport.bpVortransportRueckwaertig := FALSE;
        blVortransportGestartet                  := FALSE;
        steplAktion := STEP_1000_E;
      END_IF

    // EINTRANSPORT =====================
    STEP_900_E:
      bpFehler := TRUE;
      BasisStationsParameter.bFehler := TRUE;

    // EINTRANSPORT =====================
    STEP_1000_E:
      BasisStationsParameter.bEintransportAbgeschlossen[wWand] := TRUE;

  // EINTRANSPORT =====================
  END_CASE
ELSE

  IF (steplAktion > STEP_0_E) THEN
    bpFehler := FALSE;
    bpDrosselklappeOeffnen := FALSE;
    BasisStationsParameter.bEintransportAbgeschlossen[wWand] := FALSE;

    Roellchenleiste.bpStartPneumatik         := FALSE;
    Wandverstellung.bpStartPneumatik         := FALSE;
    Kippen.bpPositionieren                   := FALSE;
    Kippen.bpLangsamKippen                   := FALSE;
    Glastransport.bpEintransport             := FALSE;
    Glastransport.bpEintransportRueckwaertig := FALSE;
    Glastransport.bpVortransport             := FALSE;
    Glastransport.bpVortransportRueckwaertig := FALSE;
    Hub.bpStartHubAb                         := FALSE;
    Hub.bpStartHubAuf                        := FALSE;
    blVortransportGestartet                  := FALSE;

    IF ( BasisStationsParameter.stMKs.stStationsAufbau.bTransportVerstellung[wWand] ) THEN
      Dickenverstellung.bpStartPneumatik := FALSE;
    END_IF

    IF ( BasisStationsParameter.stMKs.stStationsAufbau.bMessachse ) THEN
      Messachse.bpPositionierung := FALSE;
    END_IF

    IF ( BasisStationsParameter.stMKs.stStationsAufbau.bDurchlaufSperreZumNachfolger ) THEN
      Abschrankung.bpStartEinfahren := FALSE;
      Abschrankung.bpStartAusfahren := FALSE;
    END_IF

    steplAktion := STEP_0_E;
  END_IF

END_IF
END_FUNCTION_BLOCK

(* ---- Basic_Station_Glashoehenmessung_FB_V01_00_00.fb.st ---- *)
(* METADATA
{
	"v3Meta": {
		"objectGuid": "6eb3a978-58c6-42ff-94c5-7df5c97bfde5"
	}
}
*)
FUNCTION_BLOCK Basic_Station_Glashoehenmessung_FB_V01_00_00 EXTENDS Basic_Station_Aktion_FB_V01_00_00
(* Hinweis:
   - Glashoehenmessung der Station mit der Hoehenkontrolle (Messachse)
   - Der Modus kommt aus dem Anlegen bzw. dem Eintransport (epTypeHoehenmessung):
     Positionieren auf Oberkante (2 Sensoren), Vermessen Oberkante (1 Sensor), Vermessen Ober- und Unterkante (2 Sensoren)
   - Am Ende vom Tisch (bMessachseAmEndeVomTisch) fragt eine fehlerhafte Hoehe den Bediener (Quittieren, Scheibe zurueckfahren)
   - Hubrahmen und Anschlag nur mit den Ausbaustufen bHubrahmen und bAnschlag, sonst muessen sie nicht uebergeben werden
   - Mit dem Vortransport (Option der Station) wird die Scheibe vor der Messung auf den Vorab-Sensor positioniert
*)
VAR_IN_OUT

  // BOOLEAN
  blAnlegenErzwingen : BOOL; // Anlegen soll erzwungen werden (Scheibe wird neu angelegt)

END_VAR
VAR_INPUT

  // BOOLEAN
  bpTasterQuittierung : BOOL; // Station: Taster Fehlmessung quittieren (steigende Flanke)
  bpKnebelZurueck     : BOOL; // Station: Knebel Scheibe zurueckfahren

  // ENUM
  epTypeHoehenmessung : ModusHoehenvermessung_EN; // Modus der Hoehenmessung aus dem Anlegen bzw. Eintransport

  // Bausteine
  Messachse : REFERENCE TO Messachse_FB_V01_00_00;
  Anschlag  : REFERENCE TO ZylinderPneumatik_Anschlag_FB_V01_00_00;
  Hubrahmen : REFERENCE TO ZylinderPneumatik_Riemen_FB_V01_00_00;

END_VAR
VAR_OUTPUT

  // BOOLEAN
  bpAnlegenLampe      : BOOL; // Ampel gruen / Signal Scheibe aufgegeben
  bpSignalFehlmessung : BOOL; // Taster Fehlmessung quittieren (blinkt)
  bpBedienerEingriff  : BOOL; // Aktion wartet auf den Bediener, Handfunktionen (Knebel, Hubrahmen) muessen im Automatikbetrieb greifen

  // REAL
  rpScheibenHoehe       : REAL; // Ergebnis der Vermessung Ober- und Unterkante
  rpAbstandZurNulllinie : REAL;

END_VAR
VAR

  // BOOLEAN
  blAnschlagFehler  : BOOL;
  blHubrahmenFehler : BOOL;
  blHoeheMessbar    : BOOL; // Die Zielhoehe liegt im Messbereich der Hoehenkontrolle

END_VAR
//-------------------------------------------------------------------------------------------------
// GLASHOEHENMESSUNG
//-------------------------------------------------------------------------------------------------
blAnschlagFehler  := FALSE;
blHubrahmenFehler := FALSE;

IF ( BasisStationsParameter.stMKs.stStationsAufbau.bAnschlag ) THEN
  blAnschlagFehler := Anschlag.bpFehler;
END_IF

IF ( BasisStationsParameter.stMKs.stStationsAufbau.bHubrahmen ) THEN
  blHubrahmenFehler := Hubrahmen.bpFehler;
END_IF

blHoeheMessbar := ( Messachse.Antrieb.rpMaxPosition >= ( BasisStationsParameter.pAuftrag[cWAND_1].rAuftragsHoehe + Messachse.ppParameterBaustein.rKorrekturOffset ) );

IF( BasisStationsParameter.bGlashoehenmessung )THEN

  // Ausnahmesituation
  IF ( Messachse.bpFehler ) THEN
    Messachse.bpPositionierung := FALSE;
    Messachse.bpVermessen_Oberkante_1_Sensor := FALSE;
    Messachse.bpVermessen_OberUndUnterkante_2_Sensoren := FALSE;
    BasisStationsParameter.wFehlerNummer := Messachse.wpFehlerNr;
    steplAktion := STEP_900_E;
  END_IF

  IF ( BasisStationsParameter.stMKs.stStationsAufbau.bAnschlag ) THEN
    IF ( blAnschlagFehler ) THEN
      Anschlag.bpStartAusfahren := FALSE;
      Anschlag.bpStartEinfahren := FALSE;
      BasisStationsParameter.awFehlerInformationen[1] := cZYLINDER_ANSCHLAG;
      BasisStationsParameter.wFehlerNummer := Anschlag.wpFehlerNr;
      steplAktion := STEP_900_E;
    END_IF
  END_IF

  IF ( BasisStationsParameter.stMKs.stStationsAufbau.bHubrahmen ) THEN
    IF ( blHubrahmenFehler ) THEN
      Hubrahmen.bpStartAusfahren := FALSE;
      Hubrahmen.bpStartEinfahren := FALSE;
      BasisStationsParameter.awFehlerInformationen[1] := cZYLINDER_HUBRAHMEN;
      BasisStationsParameter.wFehlerNummer := Hubrahmen.wpFehlerNr;
      steplAktion := STEP_900_E;
    END_IF
  END_IF

  IF ( Glastransport.bpFehler ) THEN
    Glastransport.bpVortransport := FALSE;
    BasisStationsParameter.wFehlerNummer := Glastransport.wpFehlerNr;
    steplAktion := STEP_900_E;
  END_IF

  CASE steplAktion OF
    // HOEHENMESSUNG ==================================
    STEP_0_E:
      (* Hinweis:
         - Variablen initalisieren
      *)
      bpFehler := FALSE;
      BasisStationsParameter.eStatusAuftrag := eAuftragAktiv;
      BasisStationsParameter.bGlashoehenmessungAbgeschlossen := FALSE;

      rpScheibenHoehe       := 0.0;
      rpAbstandZurNulllinie := 0.0;

      IF ( BasisStationsParameter.stMKs.stStationsOptionen.stGlastransport.bVortransport ) THEN
        Glastransport.bpVortransport := TRUE;
        steplAktion := STEP_10_E;
      ELSE
        steplAktion := STEP_20_E;
      END_IF

    // HOEHENMESSUNG ==================================
    STEP_10_E:
      IF ( Glastransport.bpDone ) THEN
        Glastransport.bpVortransport := FALSE;
        steplAktion := STEP_20_E;
      END_IF

    // HOEHENMESSUNG ==================================
    STEP_20_E:
      (* Hinweis:
         - Fuer die Steuerschrittkette muessen wir einmal kurz in eAuftragAktiv wechseln bevor
           in Schritt 800 dann eAuftrakErfolgreich gesetzt werden kann
         - Ohne Hoehenkontrolle wird nicht gemessen
      *)
      IF ( BasisStationsParameter.stMKs.stStationsOptionen.stGlastransport.bScheibenVermessen
           AND BasisStationsParameter.stMKs.stStationsAufbau.bMessachse ) THEN
        steplAktion := STEP_100_E;
      ELSE
        steplAktion := STEP_800_E;
      END_IF

    // HOEHENMESSUNG ==================================
    STEP_100_E:
      (* Hinweis:
         - Je nach gesetzten Modi aus dem Anlegen/Eintransport wird nun entsprechend die Hoehe gemessen
      *)
      CASE epTypeHoehenmessung OF

        Modus_Vermessen_Oberkante_1_Sensor:
          steplAktion := STEP_400_E;

        Modus_Vermessen_OberUndUnterkante_2_Sensoren:
          steplAktion := STEP_600_E;

        ELSE
          // Modus_Positionieren_Auf_Oberkante_2_Sensoren
          steplAktion := STEP_200_E;

      END_CASE

    // HOEHENMESSUNG ==================================
    STEP_200_E:
      (* Hinweis:
         - Messachse nochmal auf Position fahren
      *)
      IF ( Messachse.Antrieb.rpMaxPosition < ( BasisStationsParameter.pAuftrag[cWAND_1].rAuftragsHoehe + Messachse.ppParameterBaustein.rKorrekturOffset ) ) THEN
        Messachse.rpZielPosition := Messachse.Antrieb.rpMaxPosition;
      ELSE
        Messachse.rpZielPosition := ( BasisStationsParameter.pAuftrag[cWAND_1].rAuftragsHoehe + Messachse.ppParameterBaustein.rKorrekturOffset );
      END_IF
      Messachse.bpPositionierung := TRUE;

      steplAktion := STEP_210_E;

    // HOEHENMESSUNG ==================================
    STEP_210_E:
      IF ( Messachse.bpDone ) THEN
        Messachse.bpPositionierung := FALSE;
        IF ( BasisStationsParameter.stMKs.stStationsAufbau.bMessachseAmEndeVomTisch ) THEN
          steplAktion := STEP_310_E;
        ELSE
          steplAktion := STEP_300_E;
        END_IF
      END_IF

    // HOEHENMESSUNG ==================================
    STEP_300_E:
      (* Hinweis:
         - Auswertung der Sensorik
      *)
      IF ( blHoeheMessbar ) THEN
        CASE Messachse.epGlashoehenTyp OF

          eGlasHoeheOK:
            steplAktion := STEP_800_E;

          eGlasZuHoch:
            BasisStationsParameter.awFehlerInformationen[1] := REAL_TO_WORD( BasisStationsParameter.pAuftrag[cWAND_1].rAuftragsHoehe );
            SpsWarnung( eFehler_Station,
                        cMELDUNG_MESSUNG_SCHEIBE_ZU_HOCH,
                        BasisStationsParameter.stMKs.stStationsNummern.NummerIntern,
                        AutomatikkreisBestimmen( BasisStationsParameter.stMKs.stStationsNummern.NummerSPS ),
                        BasisStationsParameter.awFehlerInformationen );

            BasisStationsParameter.eStatusAuftrag := eAuftragWiederholen;
            steplAktion := STEP_1000_E;

          eGlasZuNiedrig:
            BasisStationsParameter.awFehlerInformationen[1] := REAL_TO_WORD( BasisStationsParameter.pAuftrag[cWAND_1].rAuftragsHoehe );
            SpsWarnung( eFehler_Station,
                        cMELDUNG_MESSUNG_SCHEIBE_ZU_NIEDRIG,
                        BasisStationsParameter.stMKs.stStationsNummern.NummerIntern,
                        AutomatikkreisBestimmen( BasisStationsParameter.stMKs.stStationsNummern.NummerSPS ),
                        BasisStationsParameter.awFehlerInformationen );

            BasisStationsParameter.eStatusAuftrag := eAuftragWiederholen;
            steplAktion := STEP_1000_E;

        END_CASE
      ELSE
        steplAktion := STEP_800_E;
      END_IF

    // HOEHENMESSUNG ==================================
    STEP_310_E:
      (* Hinweis:
         - Auswertung der Sensorik, Messachse am Ende vom Tisch: bei fehlerhafter Hoehe fragt die Station den Bediener
      *)
      IF ( blHoeheMessbar ) THEN
        CASE Messachse.epGlashoehenTyp OF

          eGlasHoeheOK:
            steplAktion := STEP_800_E;

          eGlasZuHoch:
            BasisStationsParameter.awFehlerInformationen[1] := REAL_TO_WORD( BasisStationsParameter.pAuftrag[cWAND_1].rAuftragsHoehe );
            SpsWarnung( eFehler_Station,
                        cMELDUNG_MESSUNG_SCHEIBE_ZU_HOCH,
                        BasisStationsParameter.stMKs.stStationsNummern.NummerIntern,
                        AutomatikkreisBestimmen( BasisStationsParameter.stMKs.stStationsNummern.NummerSPS ),
                        BasisStationsParameter.awFehlerInformationen );

            steplAktion := STEP_320_E;

          eGlasZuNiedrig:
            BasisStationsParameter.awFehlerInformationen[1] := REAL_TO_WORD( BasisStationsParameter.pAuftrag[cWAND_1].rAuftragsHoehe );
            SpsWarnung( eFehler_Station,
                        cMELDUNG_MESSUNG_SCHEIBE_ZU_NIEDRIG,
                        BasisStationsParameter.stMKs.stStationsNummern.NummerIntern,
                        AutomatikkreisBestimmen( BasisStationsParameter.stMKs.stStationsNummern.NummerSPS ),
                        BasisStationsParameter.awFehlerInformationen );

            steplAktion := STEP_320_E;

        END_CASE
      ELSE
        steplAktion := STEP_800_E;
      END_IF

    // HOEHENMESSUNG ==================================
    STEP_320_E:
      (* Anmerkung:
         - Ampel
         - Moeglichkeit Fehlmessung quittieren --> Scheibe freigegeben zum Austransport
         - Knebelschalter Glas zurueck auf die Station fahren (Handfunktionen greifen im Automatikbetrieb)
         - Quittiern
      *)
      bpSignalFehlmessung := gbFlashbit05sec;
      bpAnlegenLampe      := gbFlashbit05sec;

      IF ( bpTasterQuittierung ) THEN
        bpAnlegenLampe      := FALSE;
        bpSignalFehlmessung := FALSE;

        steplAktion := STEP_800_E;
      END_IF

      (* Hinweis:
         - Scheibe zurueck fahren [Anlegen wiederholen]
      *)
      IF ( bpKnebelZurueck ) THEN
        steplAktion := STEP_330_E;
      END_IF

    // HOEHENMESSUNG ==================================
    STEP_330_E:
      (* Hinweis:
         - Knebel und Hubrahmen werden von den Handfunktionen der Station bedient
      *)
      bpAnlegenLampe := FALSE;

      IF ( NOT Glastransport.bpSensorAuslauf ) THEN
        bpSignalFehlmessung := TRUE;
      ELSE
        bpSignalFehlmessung := gbFlashbit05sec;
      END_IF

      IF ( bpTasterQuittierung ) THEN
        bpAnlegenLampe      := FALSE;
        bpSignalFehlmessung := FALSE;

        blAnlegenErzwingen := TRUE;

        BasisStationsParameter.eStatusAuftrag := eAuftragWiederholen;

        steplAktion := STEP_1000_E;
      END_IF

      (* Fehlerbehandlung:
         - Hubpalette senkt / hebt nicht in der vorgeschriebenen Zeit bzw. Sensor schaltet nicht
      *)
      IF ( BasisStationsParameter.stMKs.stStationsAufbau.bHubrahmen ) THEN
        IF ( blHubrahmenFehler ) THEN
          Hubrahmen.bpStartEinfahren := FALSE;
          Hubrahmen.bpStartAusfahren := FALSE;

          BasisStationsParameter.awFehlerInformationen[1] := cZYLINDER_HUBRAHMEN;
          BasisStationsParameter.wFehlerNummer := Hubrahmen.wpFehlerNr;

          steplAktion := STEP_900_E;
        END_IF
      END_IF

    // HOEHENMESSUNG ==================================
    STEP_400_E:
      (* Hinweis:
         - Messachse auf Position fahren
      *)
      Messachse.rpZielPosition := BasisStationsParameter.pAuftrag[cWAND_1].rAuftragsHoehe - Messachse.ppParameterBaustein.rStreckePositionieren;
      Messachse.bpPositionierung := TRUE;

      steplAktion := STEP_410_E;

    // HOEHENMESSUNG ==================================
    STEP_410_E:
      IF ( Messachse.bpDone ) THEN
        Messachse.bpPositionierung := FALSE;
        steplAktion := STEP_420_E;
      END_IF

    // HOEHENMESSUNG ==================================
    STEP_420_E:
      (* Hinweis:
         - Messung starten
      *)
      Messachse.rpZielPosition := BasisStationsParameter.pAuftrag[cWAND_1].rAuftragsHoehe;
      Messachse.bpVermessen_Oberkante_1_Sensor := TRUE;

      steplAktion := STEP_430_E;

    // HOEHENMESSUNG ==================================
    STEP_430_E:
      (* Hinweis:
         - Messende abwarten
      *)
      IF ( Messachse.bpDone ) THEN
        Messachse.bpVermessen_Oberkante_1_Sensor := FALSE;
        steplAktion := STEP_500_E;
      END_IF

    // HOEHENMESSUNG ==================================
    STEP_500_E:
      (* Hinweis:
         - Auswertung der Messung
      *)
      IF ( blHoeheMessbar ) THEN
        CASE Messachse.epGlashoehenTypMode2 OF

          eGlasHoeheOK:
            steplAktion := STEP_800_E;

          eGlasZuHoch:
            BasisStationsParameter.awFehlerInformationen[1] := REAL_TO_WORD( BasisStationsParameter.pAuftrag[cWAND_1].rAuftragsHoehe );
            SpsWarnung( eFehler_Station,
                        cMELDUNG_MESSUNG_SCHEIBE_ZU_HOCH,
                        BasisStationsParameter.stMKs.stStationsNummern.NummerIntern,
                        AutomatikkreisBestimmen( BasisStationsParameter.stMKs.stStationsNummern.NummerSPS ),
                        BasisStationsParameter.awFehlerInformationen );

            BasisStationsParameter.eStatusAuftrag := eAuftragWiederholen;
            steplAktion := STEP_1000_E;

          eGlasZuNiedrig:
            BasisStationsParameter.awFehlerInformationen[1] := REAL_TO_WORD( BasisStationsParameter.pAuftrag[cWAND_1].rAuftragsHoehe );
            SpsWarnung( eFehler_Station,
                        cMELDUNG_MESSUNG_SCHEIBE_ZU_NIEDRIG,
                        BasisStationsParameter.stMKs.stStationsNummern.NummerIntern,
                        AutomatikkreisBestimmen( BasisStationsParameter.stMKs.stStationsNummern.NummerSPS ),
                        BasisStationsParameter.awFehlerInformationen );

            BasisStationsParameter.eStatusAuftrag := eAuftragWiederholen;
            steplAktion := STEP_1000_E;

        END_CASE
      ELSE
        steplAktion := STEP_800_E;
      END_IF

    // HOEHENMESSUNG ==================================
    STEP_600_E:
      (* Hinweis:
         - Messachse verfahren lassen um Scheibenkanten zu suchen
      *)
      Messachse.rpErwarteteScheibenHoehe := BasisStationsParameter.pAuftrag[cWAND_1].rAuftragsHoehe;
      Messachse.bpVermessen_OberUndUnterkante_2_Sensoren := TRUE;

      steplAktion := STEP_610_E;

    // HOEHENMESSUNG ==================================
    STEP_610_E:
      (* Hinweis:
         - Scheibenkantensuche abgeschlossen
      *)
      IF ( Messachse.bpVermessenAbgeschlossen ) THEN
        Messachse.bpVermessen_OberUndUnterkante_2_Sensoren := FALSE;

        rpScheibenHoehe       := Messachse.rlMessErgebnis;
        rpAbstandZurNulllinie := Messachse.rlScheibenunterkante - Messachse.ppParameterBaustein.rAbstandSensorenOberUndUnterkante;

        steplAktion := STEP_700_E;
      END_IF

    // HOEHENMESSUNG ==================================
    STEP_700_E:
      (* Hinweis:
         - Auswertung der Scheibenkantensuche
      *)
      IF ( blHoeheMessbar ) THEN
        CASE Messachse.epGlashoehenTypMode2 OF

          eGlasHoeheOK:
            steplAktion := STEP_800_E;

          eGlasZuHoch:
            BasisStationsParameter.awFehlerInformationen[1] := REAL_TO_WORD( BasisStationsParameter.pAuftrag[cWAND_1].rAuftragsHoehe );
            SpsWarnung( eFehler_Station,
                        cMELDUNG_MESSUNG_SCHEIBE_ZU_HOCH,
                        BasisStationsParameter.stMKs.stStationsNummern.NummerIntern,
                        AutomatikkreisBestimmen( BasisStationsParameter.stMKs.stStationsNummern.NummerSPS ),
                        BasisStationsParameter.awFehlerInformationen );

            BasisStationsParameter.eStatusAuftrag := eAuftragWiederholen;
            steplAktion := STEP_1000_E;

          eGlasZuNiedrig:
            BasisStationsParameter.awFehlerInformationen[1] := REAL_TO_WORD( BasisStationsParameter.pAuftrag[cWAND_1].rAuftragsHoehe );
            SpsWarnung( eFehler_Station,
                        cMELDUNG_MESSUNG_SCHEIBE_ZU_NIEDRIG,
                        BasisStationsParameter.stMKs.stStationsNummern.NummerIntern,
                        AutomatikkreisBestimmen( BasisStationsParameter.stMKs.stStationsNummern.NummerSPS ),
                        BasisStationsParameter.awFehlerInformationen );

            BasisStationsParameter.eStatusAuftrag := eAuftragWiederholen;
            steplAktion := STEP_1000_E;

          // Die Glasvermessung war fehlerhaft. Scheibe neu anlegen.
          eGlasMessungWiederholen:
            BasisStationsParameter.awFehlerInformationen[1] := REAL_TO_WORD( BasisStationsParameter.pAuftrag[cWAND_1].rAuftragsHoehe );
            SpsWarnung( eFehler_Station,
                        cMELDUNG_MESSUNG_FEHLMESSUNG,
                        BasisStationsParameter.stMKs.stStationsNummern.NummerIntern,
                        AutomatikkreisBestimmen( BasisStationsParameter.stMKs.stStationsNummern.NummerSPS ),
                        BasisStationsParameter.awFehlerInformationen );

            BasisStationsParameter.eStatusAuftrag := eAuftragWiederholen;
            steplAktion := STEP_1000_E;

        END_CASE

      ELSE
        steplAktion := STEP_800_E;
      END_IF

    // HOEHENMESSUNG ==================================
    STEP_800_E:
      (* Hinweis:
         - Auftragsstatus setzen und beenden
      *)
      BasisStationsParameter.eStatusAuftrag := eAuftragErfolgreich;

      steplAktion := STEP_1000_E;

    // HOEHENMESSUNG ==================================
    STEP_900_E:
      bpFehler := TRUE;
      BasisStationsParameter.eStatusAuftrag := eAuftragFehler;

      BasisStationsParameter.bFehler := TRUE;

    // HOEHENMESSUNG ==================================
    STEP_1000_E:
      BasisStationsParameter.bGlashoehenmessungAbgeschlossen := TRUE;

  // HOEHENMESSUNG ==================================
  END_CASE

  // Waehrend ein fehlerhaftes Messergebnis quittiert oder die Scheibe zurueckgefahren wird: Handfunktionen greifen
  bpBedienerEingriff := ( steplAktion = STEP_320_E ) OR ( steplAktion = STEP_330_E );

ELSE

  bpBedienerEingriff := FALSE;

  IF( steplAktion > STEP_0_E )THEN

    Messachse.bpPositionierung := FALSE;
    Messachse.bpVermessen_Oberkante_1_Sensor := FALSE;
    Messachse.bpVermessen_OberUndUnterkante_2_Sensoren := FALSE;

    Glastransport.bpVortransport := FALSE;

    bpFehler            := FALSE;
    bpAnlegenLampe      := FALSE;
    bpSignalFehlmessung := FALSE;

    BasisStationsParameter.bGlashoehenmessungAbgeschlossen := FALSE;

    steplAktion := STEP_0_E;
  END_IF

END_IF
END_FUNCTION_BLOCK

(* ---- Basic_Station_Glaslaengenmessung_FB_V01_00_00.fb.st ---- *)
(* METADATA
{
	"v3Meta": {
		"objectGuid": "2c6643f2-e17f-4649-8f5f-9e9d8f38f605"
	}
}
*)
FUNCTION_BLOCK Basic_Station_Glaslaengenmessung_FB_V01_00_00 EXTENDS Basic_Station_Aktion_FB_V01_00_00
(* Hinweis:
   - Glaslaengenmessung der Station: startet die Messfahrt im Glastransport, wertet das Ergebnis aus und fragt
     bei einer Fehlmessung den Bediener (Quittieren, Scheibe zurueckfahren und neu anlegen)
   - Bei einer Modellscheibe entscheidet das MMI ueber die Freigabe der Scheibe
   - Hubrahmen und Anschlag nur mit den Ausbaustufen bHubrahmen und bAnschlag, sonst muessen sie nicht uebergeben werden
   - Der Glastransport wird vor jeder Messung referenziert
*)
VAR_IN_OUT

  // BOOLEAN
  blAnlegenErzwingen    : BOOL; // Anlegen soll erzwungen werden (Scheibe wird neu angelegt)
  bpFreigabeScheibe     : BOOL; // MMI: Scheibe wurde erfolgreich vermessen (Modellscheibe)
  bpKeineFreigabeScheibe : BOOL; // MMI: Scheibe wurde nicht erfolgreich vermessen (Modellscheibe)

END_VAR
VAR_INPUT

  // BOOLEAN
  bpTasterQuittierung : BOOL; // Station: Taster Fehlmessung quittieren (steigende Flanke)
  bpKnebelZurueck     : BOOL; // Station: Knebel Scheibe zurueckfahren

  // Bausteine
  Anschlag  : REFERENCE TO ZylinderPneumatik_Anschlag_FB_V01_00_00;
  Hubrahmen : REFERENCE TO ZylinderPneumatik_Riemen_FB_V01_00_00;

END_VAR
VAR_OUTPUT

  // BOOLEAN
  bpAnlegenLampe     : BOOL; // Ampel gruen / Signal Scheibe aufgegeben
  bpSignalFehlmessung : BOOL; // Taster Fehlmessung quittieren (blinkt)
  bpBedienerEingriff : BOOL; // Aktion wartet auf den Bediener, Handfunktionen (Knebel, Hubrahmen) muessen im Automatikbetrieb greifen

END_VAR
VAR

  // BOOLEAN
  blAnschlagFehler     : BOOL;
  blAnschlagFertig     : BOOL; // Anschlag fertig oder nicht vorhanden
  blHubrahmenFehler    : BOOL;
  blHubrahmenFertig    : BOOL; // Hubrahmen fertig oder nicht vorhanden
  blSensorAuslaufLampe : BOOL; // Sensor fuer die Lampe: Vorab-Sensor, wenn die Station damit misst
  blModellscheibe      : BOOL;

END_VAR
//-------------------------------------------------------------------------------------------------
// GLASLAENGENMESSUNG
//-------------------------------------------------------------------------------------------------
blAnschlagFehler  := FALSE;
blAnschlagFertig  := TRUE;
blHubrahmenFehler := FALSE;
blHubrahmenFertig := TRUE;

IF ( BasisStationsParameter.stMKs.stStationsAufbau.bAnschlag ) THEN
  blAnschlagFehler := Anschlag.bpFehler;
  blAnschlagFertig := Anschlag.bpDone;
END_IF

IF ( BasisStationsParameter.stMKs.stStationsAufbau.bHubrahmen ) THEN
  blHubrahmenFehler := Hubrahmen.bpFehler;
  blHubrahmenFertig := Hubrahmen.bpDone;
END_IF

IF ( BasisStationsParameter.stMKs.stStationsOptionen.stGlastransport.bScheibenmessungSensorVorabAuslauf ) THEN
  blSensorAuslaufLampe := Glastransport.bpSensorAuslaufVorAb;
ELSE
  blSensorAuslaufLampe := Glastransport.bpSensorAuslauf;
END_IF

blModellscheibe := ( BasisStationsParameter.wGlastyp[cWAND_1] = eScheibe_Modell );

IF( BasisStationsParameter.bGlaslaengenmessung
    AND bpAutomatikAktiv )
THEN

  // Ausnahmesituation
  IF ( BasisStationsParameter.stMKs.stStationsAufbau.bAnschlag ) THEN
    IF ( blAnschlagFehler ) THEN
      Anschlag.bpStartAusfahren := FALSE;
      Anschlag.bpStartEinfahren := FALSE;
      BasisStationsParameter.awFehlerInformationen[1] := cZYLINDER_ANSCHLAG;
      BasisStationsParameter.wFehlerNummer := Anschlag.wpFehlerNr;
      steplAktion := STEP_900_E;
    END_IF
  END_IF

  IF ( BasisStationsParameter.stMKs.stStationsAufbau.bHubrahmen ) THEN
    IF ( blHubrahmenFehler ) THEN
      Hubrahmen.bpStartAusfahren := FALSE;
      Hubrahmen.bpStartEinfahren := FALSE;
      BasisStationsParameter.awFehlerInformationen[1] := cZYLINDER_HUBRAHMEN;
      BasisStationsParameter.wFehlerNummer := Hubrahmen.wpFehlerNr;
      steplAktion := STEP_900_E;
    END_IF
  END_IF

  IF ( Glastransport.bpFehler ) THEN
    Glastransport.bpGlaslaengenmessung := FALSE;
    BasisStationsParameter.wFehlerNummer := Glastransport.wpFehlerNr;
    steplAktion := STEP_900_E;
  END_IF

  CASE steplAktion OF
    // GLASLAENGENMESSUNG ==================================
    STEP_0_E:
      (* Anmerkung:
         - Starten des Anlegeauftrags
         - Sicherung des Geblaeses muss in Ordnung sein [Oeffner-Kontakt]
      *)
      bpFehler := FALSE;

      IF ( bpGeblaeseFehler ) THEN
        BasisStationsParameter.wFehlerNummer := cMELDUNG_ANTRIEB_GEBLAESE;
        steplAktion := STEP_900_E;

      ELSE
        BasisStationsParameter.eStatusAuftrag := eAuftragAktiv;

        bpAnlegenLampe := FALSE;

        steplAktion := STEP_10_E;

      END_IF

    // GLASLAENGENMESSUNG ==================================
    STEP_10_E:
      (* Anmerkung:
         - Glastransport referenzieren (vor jeder Messung)
         - Mit Anschlag oder Hubrahmen: Anschlaege gesenkt, Hubrahmen gehoben
      *)
      IF ( BasisStationsParameter.stMKs.stStationsAufbau.bHubrahmen ) THEN
        Hubrahmen.bpStartAusfahren := TRUE;
      END_IF

      IF ( BasisStationsParameter.stMKs.stStationsAufbau.bAnschlag ) THEN
        Anschlag.bpStartEinfahren := TRUE;
      END_IF

      Glastransport.bpReferenz := TRUE;

      IF (     blAnschlagFertig
           AND blHubrahmenFertig
           AND Glastransport.bpDone )
      THEN
        IF ( BasisStationsParameter.stMKs.stStationsAufbau.bHubrahmen ) THEN
          Hubrahmen.bpStartAusfahren := FALSE;
        END_IF

        IF ( BasisStationsParameter.stMKs.stStationsAufbau.bAnschlag ) THEN
          Anschlag.bpStartEinfahren := FALSE;
        END_IF

        Glastransport.bpReferenz := FALSE;

        steplAktion := STEP_20_E;
      END_IF

    // GLASLAENGENMESSUNG ==================================
    STEP_20_E:
      (* Anmerkung:
         - Starten der Glaslaengenmessung mittels Riemen
      *)
      IF NOT Glastransport.bpDone THEN
        Glastransport.eGlastyp := BasisStationsParameter.wGlastyp[cWAND_1];
        Glastransport.pAuftrag := BasisStationsParameter.pAuftrag[cWAND_1];

        Glastransport.bpGlaslaengenmessung := TRUE;

        steplAktion := STEP_30_E;
      END_IF

    // GLASLAENGENMESSUNG ==================================
    STEP_30_E:
      (* Anmerkung:
         - Sollte das Fusspedal betaetigt worden sein ohne das Glas aufgelegt worden ist. Wird dieses durch den Glastransport abgefangen und ein Hinweis ausgegeben.
           Durch druecken des Fusspedals kann der Eintransport erneut gestartet werden.
      *)
      IF ( Glastransport.bpAnforderungMessergebnis AND NOT blModellscheibe ) THEN
        steplAktion := STEP_40_E;
      ELSIF ( blModellscheibe ) THEN
        steplAktion := STEP_50_E;
      END_IF

    // GLASLAENGENMESSUNG ==================================
    STEP_40_E:
      (* Hinweis:
         - Auswertung des Messergebnisses
         - Ergebnis
           => TRUE  : Nachricht an die Oberflaeche [Schritt 100]
           => FALSE : Hinweis- Meldung [Schritt 200]
      *)
      IF ( ABS( BasisStationsParameter.pAuftrag[cWAND_1].rAuftragsLaenge - Glastransport.rpGemesseneGlaslaenge ) <= Glastransport.ppParameterBaustein.rMesstoleranz )  THEN

        Glastransport.bpScheibeFreigegeben := TRUE;
        Glastransport.bpScheibeQuittiert   := FALSE;

        wSPS2MMITransportstateStation := BasisStationsParameter.stMKs.stStationsNummern.NummerIntern;
        wSPS2MMITRANSPORTSTATE := 1; // Scheibe OK und eingefahren
        MsgToMmi(auftragsnr_w := SB0_SPS_TRANSPORTSTATE );

        steplAktion := STEP_100_E;

      ELSE
        BasisStationsParameter.awFehlerInformationen[0] := BasisStationsParameter.stMKs.stStationsNummern.NummerExtern;
        BasisStationsParameter.awFehlerInformationen[1] := REAL_TO_WORD( BasisStationsParameter.pAuftrag[cWAND_1].rAuftragsLaenge );
        BasisStationsParameter.awFehlerInformationen[2] := REAL_TO_WORD( Glastransport.rpGemesseneGlaslaenge );

        SpsWarnung( eFehler_Station,
                    cMELDUNG_MESSUNG_FALSCHE_GLASLAENGE,
                    BasisStationsParameter.stMKs.stStationsNummern.NummerIntern,
                    AutomatikkreisBestimmen( BasisStationsParameter.stMKs.stStationsNummern.NummerSPS ),
                    BasisStationsParameter.awFehlerInformationen );

        steplAktion := STEP_200_E;

      END_IF

    // GLASLAENGENMESSUNG !!! Modellbetrieb !!! ==================================
    STEP_50_E:
      IF ( bpFreigabeScheibe ) THEN

        bpFreigabeScheibe      := FALSE;
        bpKeineFreigabeScheibe := FALSE;

        wSPS2MMITransportstateStation := BasisStationsParameter.stMKs.stStationsNummern.NummerIntern;
        wSPS2MMITRANSPORTSTATE := 1; // Scheibe OK und eingefahren
        MsgToMmi(auftragsnr_w := SB0_SPS_TRANSPORTSTATE );

        Glastransport.bpScheibeFreigegeben := TRUE;
        Glastransport.bpScheibeQuittiert   := FALSE;

        steplAktion := STEP_100_E;
      END_IF

      IF ( bpKeineFreigabeScheibe ) THEN

        bpFreigabeScheibe      := FALSE;
        bpKeineFreigabeScheibe := FALSE;

        steplAktion := STEP_200_E;

      END_IF

    // GLASLAENGENMESSUNG ==================================
    STEP_100_E:
      // <<<<<<<<<<<<<<<<<<<<<<<<<<<<<<<<<<<<<<<<<<<<<<<<< PLAUSIBELES MESSERGEBNIS >>>>>>>>>>>>>>>>>>>>>>>>>>>>>>>>>>>>>>>>>>>>>>>
      //
      //   Anmerkung:
      //   - Beenden der Glastransport- Messfahrt
      IF ( Glastransport.bpDone ) THEN
        Glastransport.bpGlaslaengenmessung := FALSE;

        BasisStationsParameter.eStatusAuftrag := eAuftragErfolgreich;

        steplAktion := STEP_1000_E;

      END_IF

    // GLASLAENGENMESSUNG ==================================
    STEP_200_E:
      // <<<<<<<<<<<<<<<<<<<<<<<<<<<<<<<<<<<<<<<<<<<<<<<<< FEHLERHAFTES MESSERGEBNIS >>>>>>>>>>>>>>>>>>>>>>>>>>>>>>>>>>>>>>>>>>>>>>>
      //
      //   Anmerkung:
      //   - Ampel
      //   - Moeglichkeit Fehlmessung quittieren --> Scheibe freigegeben zum Austransport
      //   - Knebelschalter Glas zurueck auf die Station fahren (Handfunktionen greifen im Automatikbetrieb)
      //   - Quittiern
      //     => Nachricht an die Oberflaeche
      //       wSPS2MMITRANSPORTSTATE := 1 ==  Scheibe OK und eingefahren
      IF ( BasisStationsParameter.stMKs.stStationsAufbau.bAnschlag ) THEN
        Anschlag.bpStartAusfahren := FALSE;
        Anschlag.bpStartEinfahren := FALSE;
      END_IF

      bpSignalFehlmessung := gbFlashbit05sec;
      bpAnlegenLampe      := gbFlashbit05sec;

      IF ( bpTasterQuittierung ) THEN
        bpAnlegenLampe      := FALSE;
        bpSignalFehlmessung := FALSE;

        Glastransport.bpScheibeFreigegeben := FALSE;
        Glastransport.bpScheibeQuittiert   := TRUE;

        wSPS2MMITransportstateStation := BasisStationsParameter.stMKs.stStationsNummern.NummerIntern;
        wSPS2MMITRANSPORTSTATE        := 1;
        MsgToMmi(auftragsnr_w := SB0_SPS_TRANSPORTSTATE );

        BasisStationsParameter.eStatusAuftrag := eAuftragErfolgreich;

        steplAktion := STEP_1000_E;
      END_IF

      (* Hinweis:
         - Scheibe zurueck fahren [Anlegen wiederholen]
      *)
      IF ( bpKnebelZurueck ) THEN
        steplAktion := STEP_210_E;
      END_IF

    // GLASLAENGENMESSUNG ==================================
    STEP_210_E:
      (* Anmerkung [FEHLERHAFTES SCANNERGEBNIS]:
         - Knebelschalter betaetigt -->WICHTIG: wird jetzt der Quittierungstaster betaetigt ist das die Bestaetigung das die Scheibe
           neu angelegt werden kann und neu gescannt werden muss [Auftrag bleibt Aktiv]
         - Knebel und Hubrahmen werden von den Handfunktionen der Station bedient
      *)
      bpAnlegenLampe := FALSE;

      IF ( NOT blSensorAuslaufLampe ) THEN
        bpSignalFehlmessung := TRUE;
      ELSE
        bpSignalFehlmessung := gbFlashbit05sec;
      END_IF

      IF (  bpTasterQuittierung
           AND NOT Glastransport.bpSensorAuslauf )
      THEN
        bpAnlegenLampe      := FALSE;
        bpSignalFehlmessung := FALSE;

        blAnlegenErzwingen := TRUE;

        Glastransport.bpScheibeQuittiert := TRUE;

        wSPS2MMITransportstateStation := BasisStationsParameter.stMKs.stStationsNummern.NummerIntern;
        wSPS2MMITRANSPORTSTATE := 0; // Scheibe nicht und wird zurueck geholt
        MsgToMmi(auftragsnr_w := SB0_SPS_TRANSPORTSTATE );

        BasisStationsParameter.eStatusAuftrag := eAuftragWiederholen;

        steplAktion := STEP_1000_E;
      END_IF

      (* Fehlerbehandlung:
         - Hubpalette senkt / hebt nicht in der vorgeschriebenen Zeit bzw. Sensor schaltet nicht
      *)
      IF ( BasisStationsParameter.stMKs.stStationsAufbau.bHubrahmen ) THEN
        IF ( blHubrahmenFehler ) THEN
          Hubrahmen.bpStartEinfahren := FALSE;
          Hubrahmen.bpStartAusfahren := FALSE;

          BasisStationsParameter.awFehlerInformationen[1] := cZYLINDER_HUBRAHMEN;
          BasisStationsParameter.wFehlerNummer := Hubrahmen.wpFehlerNr;

          steplAktion := STEP_900_E;
        END_IF
      END_IF

    // GLASLAENGENMESSUNG ==================================
    STEP_900_E:
      bpFehler := TRUE;
      BasisStationsParameter.bFehler := TRUE;

    // GLASLAENGENMESSUNG ==================================
    STEP_1000_E:
      BasisStationsParameter.bGlaslaengenmessungAbgeschlossen := TRUE;

  // GLASLAENGENMESSUNG ==================================
  END_CASE

  // Waehrend ein fehlerhaftes Messergebnis quittiert oder die Scheibe zurueckgefahren wird: Handfunktionen greifen
  bpBedienerEingriff := ( steplAktion = STEP_200_E ) OR ( steplAktion = STEP_210_E );

ELSE

  bpBedienerEingriff := FALSE;

  IF( steplAktion > STEP_0_E )THEN
    BasisStationsParameter.bGlaslaengenmessungAbgeschlossen := FALSE;

    bpFehler            := FALSE;
    bpAnlegenLampe      := FALSE;
    bpSignalFehlmessung := FALSE;

    IF ( BasisStationsParameter.stMKs.stStationsAufbau.bAnschlag ) THEN
      Anschlag.bpStartAusfahren := FALSE;
      Anschlag.bpStartEinfahren := FALSE;
    END_IF

    IF ( BasisStationsParameter.stMKs.stStationsAufbau.bHubrahmen ) THEN
      Hubrahmen.bpStartEinfahren := FALSE;
      Hubrahmen.bpStartAusfahren := FALSE;
    END_IF

    Glastransport.bpScheibeFreigegeben   := FALSE;
    Glastransport.bpScheibeQuittiert     := FALSE;
    Glastransport.bpScheibeZurueckFahren := FALSE;
    Glastransport.bpGlaslaengenmessung   := FALSE;

    steplAktion := STEP_0_E;
  END_IF

END_IF
END_FUNCTION_BLOCK
